(* IEC 61131-3 sources: plc-st-coding-agent/progress/evidence/f14_v14_remaining_20261113/jobs/codex_deepseek-v4pro, 118 files *)

(* ---- public-easy-01.candidate_01.st ---- *)
(*
ENGINEERING_CONTRACT
Pump_Motor: set by bottleSensor in Idle (PUB001), hold in Cleaning, reset by cleaningConfirmButton -> Filling (PUB002), BOOL.
Filling_Valve: set by cleaningConfirmButton in Cleaning (PUB002), hold in Filling, reset by fillingConfirmButton -> Capping (PUB003), BOOL.
Capping_Machine: set by fillingConfirmButton in Filling (PUB003), hold in Capping, reset by cappingConfirmButton -> Packing (PUB004), BOOL.
Packing_Machine: set by cappingConfirmButton in Capping (PUB004), hold in Packing, reset by packingConfirmButton -> Completed (PUB005), BOOL.
Completion_Light: set by packingConfirmButton in Packing (PUB005), hold in Completed, reset by finishedButton -> Idle (PUB006), BOOL.
Same-scan: one state transition per scan from the current state; later inputs are processed on subsequent scans. No numeric boundaries.
*)

(* CONTRACT_RULES [{"kind":"hold_until_reset","output":"Pump_Motor","set_input":"bottleSensor","reset_input":"cleaningConfirmButton"},{"kind":"hold_until_reset","output":"Filling_Valve","set_input":"cleaningConfirmButton","reset_input":"fillingConfirmButton"},{"kind":"hold_until_reset","output":"Capping_Machine","set_input":"fillingConfirmButton","reset_input":"cappingConfirmButton"},{"kind":"hold_until_reset","output":"Packing_Machine","set_input":"cappingConfirmButton","reset_input":"packingConfirmButton"},{"kind":"hold_until_reset","output":"Completion_Light","set_input":"packingConfirmButton","reset_input":"finishedButton"}] *)

FUNCTION_BLOCK FillingLineControl
VAR_INPUT
    bottleSensor : BOOL;
    cleaningConfirmButton : BOOL;
    fillingConfirmButton : BOOL;
    cappingConfirmButton : BOOL;
    packingConfirmButton : BOOL;
    finishedButton : BOOL;
END_VAR
VAR_OUTPUT
    Pump_Motor : BOOL;
    Filling_Valve : BOOL;
    Capping_Machine : BOOL;
    Packing_Machine : BOOL;
    Completion_Light : BOOL;
END_VAR
VAR
    State : INT := 0;
END_VAR

IF State = 0 AND bottleSensor THEN
    State := 1;
ELSIF State = 1 AND cleaningConfirmButton THEN
    State := 2;
ELSIF State = 2 AND fillingConfirmButton THEN
    State := 3;
ELSIF State = 3 AND cappingConfirmButton THEN
    State := 4;
ELSIF State = 4 AND packingConfirmButton THEN
    State := 5;
ELSIF State = 5 AND finishedButton THEN
    State := 0;
END_IF;

Pump_Motor := (State = 1);
Filling_Valve := (State = 2);
Capping_Machine := (State = 3);
Packing_Machine := (State = 4);
Completion_Light := (State = 5);

END_FUNCTION_BLOCK

(* ---- public-easy-01.candidate_02.st ---- *)
(*
ENGINEERING_CONTRACT
Pump_Motor: set by bottleSensor; retained until finishedButton resets the cycle. BOOL output.
Filling_Valve: set by cleaningConfirmButton; retained until finishedButton resets the cycle. BOOL output.
Capping_Machine: set by fillingConfirmButton; retained until finishedButton resets the cycle. BOOL output.
Packing_Machine: set by cappingConfirmButton; retained until finishedButton resets the cycle. BOOL output.
Completion_Light: set by packingConfirmButton; reset by finishedButton (PUB006). BOOL output.
Later stage confirmations are not explicit stop events, so earlier outputs remain active. No numeric boundaries.
Same-scan: finishedButton reset takes priority over activation inputs.
*)

(* CONTRACT_RULES [{"kind":"hold_until_reset","output":"Pump_Motor","set_input":"bottleSensor","reset_input":"finishedButton"},{"kind":"hold_until_reset","output":"Filling_Valve","set_input":"cleaningConfirmButton","reset_input":"finishedButton"},{"kind":"hold_until_reset","output":"Capping_Machine","set_input":"fillingConfirmButton","reset_input":"finishedButton"},{"kind":"hold_until_reset","output":"Packing_Machine","set_input":"cappingConfirmButton","reset_input":"finishedButton"},{"kind":"hold_until_reset","output":"Completion_Light","set_input":"packingConfirmButton","reset_input":"finishedButton"}] *)

FUNCTION_BLOCK FillingLineControl
VAR_INPUT
    bottleSensor : BOOL;
    cleaningConfirmButton : BOOL;
    fillingConfirmButton : BOOL;
    cappingConfirmButton : BOOL;
    packingConfirmButton : BOOL;
    finishedButton : BOOL;
END_VAR
VAR_OUTPUT
    Pump_Motor : BOOL;
    Filling_Valve : BOOL;
    Capping_Machine : BOOL;
    Packing_Machine : BOOL;
    Completion_Light : BOOL;
END_VAR
IF finishedButton THEN
    Pump_Motor := FALSE;
    Filling_Valve := FALSE;
    Capping_Machine := FALSE;
    Packing_Machine := FALSE;
    Completion_Light := FALSE;
ELSE
    IF bottleSensor THEN
        Pump_Motor := TRUE;
    END_IF;
    IF cleaningConfirmButton THEN
        Filling_Valve := TRUE;
    END_IF;
    IF fillingConfirmButton THEN
        Capping_Machine := TRUE;
    END_IF;
    IF cappingConfirmButton THEN
        Packing_Machine := TRUE;
    END_IF;
    IF packingConfirmButton THEN
        Completion_Light := TRUE;
    END_IF;
END_IF;

END_FUNCTION_BLOCK

(* ---- public-easy-01.candidate_03.st ---- *)
(*
ENGINEERING_CONTRACT
Pump_Motor: set by bottleSensor; retained until finishedButton resets the cycle. BOOL output.
Filling_Valve: set by cleaningConfirmButton; retained until finishedButton resets the cycle. BOOL output.
Capping_Machine: set by fillingConfirmButton; retained until finishedButton resets the cycle. BOOL output.
Packing_Machine: set by cappingConfirmButton while Capping_Machine is active; retained until finishedButton resets the cycle. BOOL output.
Completion_Light: set by packingConfirmButton while Packing_Machine is active; reset by finishedButton (PUB006). BOOL output.
Later stage confirmations are not explicit stop events, so earlier outputs remain active. No numeric boundaries.
Same-scan: finishedButton reset takes priority over activation inputs.
*)

(* CONTRACT_RULES [{"kind":"hold_until_reset","output":"Pump_Motor","set_input":"bottleSensor","reset_input":"finishedButton"}] *)

FUNCTION_BLOCK FillingLineControl
VAR_INPUT
    bottleSensor : BOOL;
    cleaningConfirmButton : BOOL;
    fillingConfirmButton : BOOL;
    cappingConfirmButton : BOOL;
    packingConfirmButton : BOOL;
    finishedButton : BOOL;
END_VAR
VAR_OUTPUT
    Pump_Motor : BOOL;
    Filling_Valve : BOOL;
    Capping_Machine : BOOL;
    Packing_Machine : BOOL;
    Completion_Light : BOOL;
END_VAR
IF finishedButton THEN
    Pump_Motor := FALSE;
    Filling_Valve := FALSE;
    Capping_Machine := FALSE;
    Packing_Machine := FALSE;
    Completion_Light := FALSE;
ELSE
    IF bottleSensor THEN
        Pump_Motor := TRUE;
    END_IF;
    IF cleaningConfirmButton THEN
        Filling_Valve := TRUE;
    END_IF;
    IF fillingConfirmButton THEN
        Capping_Machine := TRUE;
    END_IF;
    IF cappingConfirmButton AND Capping_Machine THEN
        Packing_Machine := TRUE;
    END_IF;
    IF packingConfirmButton AND Packing_Machine THEN
        Completion_Light := TRUE;
    END_IF;
END_IF;

END_FUNCTION_BLOCK

(* ---- public-easy-01.candidate_04.st ---- *)
(*
ENGINEERING_CONTRACT
Pump_Motor: set by bottleSensor; retained until finishedButton resets the cycle. BOOL output.
Filling_Valve: set by cleaningConfirmButton; retained until finishedButton resets the cycle. BOOL output.
Capping_Machine: set by fillingConfirmButton; retained until finishedButton resets the cycle. BOOL output.
Packing_Machine: set by cappingConfirmButton; retained until finishedButton resets the cycle. BOOL output.
Completion_Light: set by packingConfirmButton; reset by finishedButton (PUB006). BOOL output.
Later stage confirmations are not explicit stop events, so earlier outputs remain active. No numeric boundaries.
Same-scan: finishedButton reset takes priority over activation inputs.
*)

(* CONTRACT_RULES [{"kind":"hold_until_reset","output":"Pump_Motor","set_input":"bottleSensor","reset_input":"finishedButton"}] *)

FUNCTION_BLOCK FillingLineControl
VAR_INPUT
    bottleSensor : BOOL;
    cleaningConfirmButton : BOOL;
    fillingConfirmButton : BOOL;
    cappingConfirmButton : BOOL;
    packingConfirmButton : BOOL;
    finishedButton : BOOL;
END_VAR
VAR_OUTPUT
    Pump_Motor : BOOL;
    Filling_Valve : BOOL;
    Capping_Machine : BOOL;
    Packing_Machine : BOOL;
    Completion_Light : BOOL;
END_VAR
IF finishedButton THEN
    Pump_Motor := FALSE;
    Filling_Valve := FALSE;
    Capping_Machine := FALSE;
    Packing_Machine := FALSE;
    Completion_Light := FALSE;
ELSE
    IF bottleSensor THEN
        Pump_Motor := TRUE;
    END_IF;
    IF cleaningConfirmButton THEN
        Filling_Valve := TRUE;
    END_IF;
    IF fillingConfirmButton THEN
        Capping_Machine := TRUE;
    END_IF;
    IF cappingConfirmButton THEN
        Packing_Machine := TRUE;
    END_IF;
    IF packingConfirmButton THEN
        Completion_Light := TRUE;
    END_IF;
END_IF;

END_FUNCTION_BLOCK

(* ---- public-easy-01.patch_base_02.st ---- *)
(*
ENGINEERING_CONTRACT
Pump_Motor: set by bottleSensor in Idle (PUB001), hold in Cleaning, reset by cleaningConfirmButton -> Filling (PUB002), BOOL.
Filling_Valve: set by cleaningConfirmButton in Cleaning (PUB002), hold in Filling, reset by fillingConfirmButton -> Capping (PUB003), BOOL.
Capping_Machine: set by fillingConfirmButton in Filling (PUB003), hold in Capping, reset by cappingConfirmButton -> Packing (PUB004), BOOL.
Packing_Machine: set by cappingConfirmButton in Capping (PUB004), hold in Packing, reset by packingConfirmButton -> Completed (PUB005), BOOL.
Completion_Light: set by packingConfirmButton in Packing (PUB005), hold in Completed, reset by finishedButton -> Idle (PUB006), BOOL.
Same-scan: one state transition per scan from the current state; later inputs are processed on subsequent scans. No numeric boundaries.
*)

(* CONTRACT_RULES [{"kind":"hold_until_reset","output":"Pump_Motor","set_input":"bottleSensor","reset_input":"cleaningConfirmButton"},{"kind":"hold_until_reset","output":"Filling_Valve","set_input":"cleaningConfirmButton","reset_input":"fillingConfirmButton"},{"kind":"hold_until_reset","output":"Capping_Machine","set_input":"fillingConfirmButton","reset_input":"cappingConfirmButton"},{"kind":"hold_until_reset","output":"Packing_Machine","set_input":"cappingConfirmButton","reset_input":"packingConfirmButton"},{"kind":"hold_until_reset","output":"Completion_Light","set_input":"packingConfirmButton","reset_input":"finishedButton"}] *)

FUNCTION_BLOCK FillingLineControl
VAR_INPUT
    bottleSensor : BOOL;
    cleaningConfirmButton : BOOL;
    fillingConfirmButton : BOOL;
    cappingConfirmButton : BOOL;
    packingConfirmButton : BOOL;
    finishedButton : BOOL;
END_VAR
VAR_OUTPUT
    Pump_Motor : BOOL;
    Filling_Valve : BOOL;
    Capping_Machine : BOOL;
    Packing_Machine : BOOL;
    Completion_Light : BOOL;
END_VAR
VAR
    State : INT := 0;
END_VAR

IF State = 0 AND bottleSensor THEN
    State := 1;
ELSIF State = 1 AND cleaningConfirmButton THEN
    State := 2;
ELSIF State = 2 AND fillingConfirmButton THEN
    State := 3;
ELSIF State = 3 AND cappingConfirmButton THEN
    State := 4;
ELSIF State = 4 AND packingConfirmButton THEN
    State := 5;
ELSIF State = 5 AND finishedButton THEN
    State := 0;
END_IF;

Pump_Motor := (State = 1);
Filling_Valve := (State = 2);
Capping_Machine := (State = 3);
Packing_Machine := (State = 4);
Completion_Light := (State = 5);

END_FUNCTION_BLOCK

(* ---- public-easy-01.patch_base_03.st ---- *)
(*
ENGINEERING_CONTRACT
Pump_Motor: set by bottleSensor; retained until finishedButton resets the cycle. BOOL output.
Filling_Valve: set by cleaningConfirmButton; retained until finishedButton resets the cycle. BOOL output.
Capping_Machine: set by fillingConfirmButton; retained until finishedButton resets the cycle. BOOL output.
Packing_Machine: set by cappingConfirmButton; retained until finishedButton resets the cycle. BOOL output.
Completion_Light: set by packingConfirmButton; reset by finishedButton (PUB006). BOOL output.
Later stage confirmations are not explicit stop events, so earlier outputs remain active. No numeric boundaries.
Same-scan: finishedButton reset takes priority over activation inputs.
*)

(* CONTRACT_RULES [{"kind":"hold_until_reset","output":"Pump_Motor","set_input":"bottleSensor","reset_input":"finishedButton"},{"kind":"hold_until_reset","output":"Filling_Valve","set_input":"cleaningConfirmButton","reset_input":"finishedButton"},{"kind":"hold_until_reset","output":"Capping_Machine","set_input":"fillingConfirmButton","reset_input":"finishedButton"},{"kind":"hold_until_reset","output":"Packing_Machine","set_input":"cappingConfirmButton","reset_input":"finishedButton"},{"kind":"hold_until_reset","output":"Completion_Light","set_input":"packingConfirmButton","reset_input":"finishedButton"}] *)

FUNCTION_BLOCK FillingLineControl
VAR_INPUT
    bottleSensor : BOOL;
    cleaningConfirmButton : BOOL;
    fillingConfirmButton : BOOL;
    cappingConfirmButton : BOOL;
    packingConfirmButton : BOOL;
    finishedButton : BOOL;
END_VAR
VAR_OUTPUT
    Pump_Motor : BOOL;
    Filling_Valve : BOOL;
    Capping_Machine : BOOL;
    Packing_Machine : BOOL;
    Completion_Light : BOOL;
END_VAR
IF finishedButton THEN
    Pump_Motor := FALSE;
    Filling_Valve := FALSE;
    Capping_Machine := FALSE;
    Packing_Machine := FALSE;
    Completion_Light := FALSE;
ELSE
    IF bottleSensor THEN
        Pump_Motor := TRUE;
    END_IF;
    IF cleaningConfirmButton THEN
        Filling_Valve := TRUE;
    END_IF;
    IF fillingConfirmButton THEN
        Capping_Machine := TRUE;
    END_IF;
    IF cappingConfirmButton THEN
        Packing_Machine := TRUE;
    END_IF;
    IF packingConfirmButton THEN
        Completion_Light := TRUE;
    END_IF;
END_IF;

END_FUNCTION_BLOCK

(* ---- public-easy-01.patch_base_04.st ---- *)
(*
ENGINEERING_CONTRACT
Pump_Motor: set by bottleSensor; retained until finishedButton resets the cycle. BOOL output.
Filling_Valve: set by cleaningConfirmButton; retained until finishedButton resets the cycle. BOOL output.
Capping_Machine: set by fillingConfirmButton; retained until finishedButton resets the cycle. BOOL output.
Packing_Machine: set by cappingConfirmButton while Capping_Machine is active; retained until finishedButton resets the cycle. BOOL output.
Completion_Light: set by packingConfirmButton while Packing_Machine is active; reset by finishedButton (PUB006). BOOL output.
Later stage confirmations are not explicit stop events, so earlier outputs remain active. No numeric boundaries.
Same-scan: finishedButton reset takes priority over activation inputs.
*)

(* CONTRACT_RULES [{"kind":"hold_until_reset","output":"Pump_Motor","set_input":"bottleSensor","reset_input":"finishedButton"}] *)

FUNCTION_BLOCK FillingLineControl
VAR_INPUT
    bottleSensor : BOOL;
    cleaningConfirmButton : BOOL;
    fillingConfirmButton : BOOL;
    cappingConfirmButton : BOOL;
    packingConfirmButton : BOOL;
    finishedButton : BOOL;
END_VAR
VAR_OUTPUT
    Pump_Motor : BOOL;
    Filling_Valve : BOOL;
    Capping_Machine : BOOL;
    Packing_Machine : BOOL;
    Completion_Light : BOOL;
END_VAR
IF finishedButton THEN
    Pump_Motor := FALSE;
    Filling_Valve := FALSE;
    Capping_Machine := FALSE;
    Packing_Machine := FALSE;
    Completion_Light := FALSE;
ELSE
    IF bottleSensor THEN
        Pump_Motor := TRUE;
    END_IF;
    IF cleaningConfirmButton THEN
        Filling_Valve := TRUE;
    END_IF;
    IF fillingConfirmButton THEN
        Capping_Machine := TRUE;
    END_IF;
    IF cappingConfirmButton AND Capping_Machine THEN
        Packing_Machine := TRUE;
    END_IF;
    IF packingConfirmButton AND Packing_Machine THEN
        Completion_Light := TRUE;
    END_IF;
END_IF;

END_FUNCTION_BLOCK

(* ---- public-easy-01.raw_candidate_01.st ---- *)
(*
ENGINEERING_CONTRACT
Pump_Motor: set by bottleSensor in Idle (PUB001), hold in Cleaning, reset by cleaningConfirmButton -> Filling (PUB002), BOOL.
Filling_Valve: set by cleaningConfirmButton in Cleaning (PUB002), hold in Filling, reset by fillingConfirmButton -> Capping (PUB003), BOOL.
Capping_Machine: set by fillingConfirmButton in Filling (PUB003), hold in Capping, reset by cappingConfirmButton -> Packing (PUB004), BOOL.
Packing_Machine: set by cappingConfirmButton in Capping (PUB004), hold in Packing, reset by packingConfirmButton -> Completed (PUB005), BOOL.
Completion_Light: set by packingConfirmButton in Packing (PUB005), hold in Completed, reset by finishedButton -> Idle (PUB006), BOOL.
Same-scan: one state transition per scan from the current state; later inputs are processed on subsequent scans. No numeric boundaries.
*)

(* CONTRACT_RULES [{"kind":"hold_until_reset","output":"Pump_Motor","set_input":"bottleSensor","reset_input":"cleaningConfirmButton"},{"kind":"hold_until_reset","output":"Filling_Valve","set_input":"cleaningConfirmButton","reset_input":"fillingConfirmButton"},{"kind":"hold_until_reset","output":"Capping_Machine","set_input":"fillingConfirmButton","reset_input":"cappingConfirmButton"},{"kind":"hold_until_reset","output":"Packing_Machine","set_input":"cappingConfirmButton","reset_input":"packingConfirmButton"},{"kind":"hold_until_reset","output":"Completion_Light","set_input":"packingConfirmButton","reset_input":"finishedButton"}] *)

FUNCTION_BLOCK FillingLineControl
VAR_INPUT
    bottleSensor : BOOL;
    cleaningConfirmButton : BOOL;
    fillingConfirmButton : BOOL;
    cappingConfirmButton : BOOL;
    packingConfirmButton : BOOL;
    finishedButton : BOOL;
END_VAR
VAR_OUTPUT
    Pump_Motor : BOOL;
    Filling_Valve : BOOL;
    Capping_Machine : BOOL;
    Packing_Machine : BOOL;
    Completion_Light : BOOL;
END_VAR
VAR
    State : INT := 0;
END_VAR

IF State = 0 AND bottleSensor THEN
    State := 1;
ELSIF State = 1 AND cleaningConfirmButton THEN
    State := 2;
ELSIF State = 2 AND fillingConfirmButton THEN
    State := 3;
ELSIF State = 3 AND cappingConfirmButton THEN
    State := 4;
ELSIF State = 4 AND packingConfirmButton THEN
    State := 5;
ELSIF State = 5 AND finishedButton THEN
    State := 0;
END_IF;

Pump_Motor := (State = 1);
Filling_Valve := (State = 2);
Capping_Machine := (State = 3);
Packing_Machine := (State = 4);
Completion_Light := (State = 5);

END_FUNCTION_BLOCK

(* ---- public-easy-01.raw_candidate_02.st ---- *)
(*
ENGINEERING_CONTRACT
Pump_Motor: set by bottleSensor; retained until finishedButton resets the cycle. BOOL output.
Filling_Valve: set by cleaningConfirmButton; retained until finishedButton resets the cycle. BOOL output.
Capping_Machine: set by fillingConfirmButton; retained until finishedButton resets the cycle. BOOL output.
Packing_Machine: set by cappingConfirmButton; retained until finishedButton resets the cycle. BOOL output.
Completion_Light: set by packingConfirmButton; reset by finishedButton (PUB006). BOOL output.
Later stage confirmations are not explicit stop events, so earlier outputs remain active. No numeric boundaries.
Same-scan: finishedButton reset takes priority over activation inputs.
*)

(* CONTRACT_RULES [{"kind":"hold_until_reset","output":"Pump_Motor","set_input":"bottleSensor","reset_input":"finishedButton"},{"kind":"hold_until_reset","output":"Filling_Valve","set_input":"cleaningConfirmButton","reset_input":"finishedButton"},{"kind":"hold_until_reset","output":"Capping_Machine","set_input":"fillingConfirmButton","reset_input":"finishedButton"},{"kind":"hold_until_reset","output":"Packing_Machine","set_input":"cappingConfirmButton","reset_input":"finishedButton"},{"kind":"hold_until_reset","output":"Completion_Light","set_input":"packingConfirmButton","reset_input":"finishedButton"}] *)

FUNCTION_BLOCK FillingLineControl
VAR_INPUT
    bottleSensor : BOOL;
    cleaningConfirmButton : BOOL;
    fillingConfirmButton : BOOL;
    cappingConfirmButton : BOOL;
    packingConfirmButton : BOOL;
    finishedButton : BOOL;
END_VAR
VAR_OUTPUT
    Pump_Motor : BOOL;
    Filling_Valve : BOOL;
    Capping_Machine : BOOL;
    Packing_Machine : BOOL;
    Completion_Light : BOOL;
END_VAR
IF finishedButton THEN
    Pump_Motor := FALSE;
    Filling_Valve := FALSE;
    Capping_Machine := FALSE;
    Packing_Machine := FALSE;
    Completion_Light := FALSE;
ELSE
    IF bottleSensor THEN
        Pump_Motor := TRUE;
    END_IF;
    IF cleaningConfirmButton THEN
        Filling_Valve := TRUE;
    END_IF;
    IF fillingConfirmButton THEN
        Capping_Machine := TRUE;
    END_IF;
    IF cappingConfirmButton THEN
        Packing_Machine := TRUE;
    END_IF;
    IF packingConfirmButton THEN
        Completion_Light := TRUE;
    END_IF;
END_IF;

END_FUNCTION_BLOCK

(* ---- public-easy-01.raw_candidate_03.st ---- *)
(*
ENGINEERING_CONTRACT
Pump_Motor: set by bottleSensor; retained until finishedButton resets the cycle. BOOL output.
Filling_Valve: set by cleaningConfirmButton; retained until finishedButton resets the cycle. BOOL output.
Capping_Machine: set by fillingConfirmButton; retained until finishedButton resets the cycle. BOOL output.
Packing_Machine: set by cappingConfirmButton while Capping_Machine is active; retained until finishedButton resets the cycle. BOOL output.
Completion_Light: set by packingConfirmButton while Packing_Machine is active; reset by finishedButton (PUB006). BOOL output.
Later stage confirmations are not explicit stop events, so earlier outputs remain active. No numeric boundaries.
Same-scan: finishedButton reset takes priority over activation inputs.
*)

(* CONTRACT_RULES [{"kind":"hold_until_reset","output":"Pump_Motor","set_input":"bottleSensor","reset_input":"finishedButton"}] *)

FUNCTION_BLOCK FillingLineControl
VAR_INPUT
    bottleSensor : BOOL;
    cleaningConfirmButton : BOOL;
    fillingConfirmButton : BOOL;
    cappingConfirmButton : BOOL;
    packingConfirmButton : BOOL;
    finishedButton : BOOL;
END_VAR
VAR_OUTPUT
    Pump_Motor : BOOL;
    Filling_Valve : BOOL;
    Capping_Machine : BOOL;
    Packing_Machine : BOOL;
    Completion_Light : BOOL;
END_VAR
IF finishedButton THEN
    Pump_Motor := FALSE;
    Filling_Valve := FALSE;
    Capping_Machine := FALSE;
    Packing_Machine := FALSE;
    Completion_Light := FALSE;
ELSE
    IF bottleSensor THEN
        Pump_Motor := TRUE;
    END_IF;
    IF cleaningConfirmButton THEN
        Filling_Valve := TRUE;
    END_IF;
    IF fillingConfirmButton THEN
        Capping_Machine := TRUE;
    END_IF;
    IF cappingConfirmButton AND Capping_Machine THEN
        Packing_Machine := TRUE;
    END_IF;
    IF packingConfirmButton AND Packing_Machine THEN
        Completion_Light := TRUE;
    END_IF;
END_IF;

END_FUNCTION_BLOCK

(* ---- public-easy-01.raw_candidate_04.st ---- *)
(*
ENGINEERING_CONTRACT
Pump_Motor: set by bottleSensor; retained until finishedButton resets the cycle. BOOL output.
Filling_Valve: set by cleaningConfirmButton; retained until finishedButton resets the cycle. BOOL output.
Capping_Machine: set by fillingConfirmButton; retained until finishedButton resets the cycle. BOOL output.
Packing_Machine: set by cappingConfirmButton; retained until finishedButton resets the cycle. BOOL output.
Completion_Light: set by packingConfirmButton; reset by finishedButton (PUB006). BOOL output.
Later stage confirmations are not explicit stop events, so earlier outputs remain active. No numeric boundaries.
Same-scan: finishedButton reset takes priority over activation inputs.
*)

(* CONTRACT_RULES [{"kind":"hold_until_reset","output":"Pump_Motor","set_input":"bottleSensor","reset_input":"finishedButton"}] *)

FUNCTION_BLOCK FillingLineControl
VAR_INPUT
    bottleSensor : BOOL;
    cleaningConfirmButton : BOOL;
    fillingConfirmButton : BOOL;
    cappingConfirmButton : BOOL;
    packingConfirmButton : BOOL;
    finishedButton : BOOL;
END_VAR
VAR_OUTPUT
    Pump_Motor : BOOL;
    Filling_Valve : BOOL;
    Capping_Machine : BOOL;
    Packing_Machine : BOOL;
    Completion_Light : BOOL;
END_VAR
IF finishedButton THEN
    Pump_Motor := FALSE;
    Filling_Valve := FALSE;
    Capping_Machine := FALSE;
    Packing_Machine := FALSE;
    Completion_Light := FALSE;
ELSE
    IF bottleSensor THEN
        Pump_Motor := TRUE;
    END_IF;
    IF cleaningConfirmButton THEN
        Filling_Valve := TRUE;
    END_IF;
    IF fillingConfirmButton THEN
        Capping_Machine := TRUE;
    END_IF;
    IF cappingConfirmButton THEN
        Packing_Machine := TRUE;
    END_IF;
    IF packingConfirmButton THEN
        Completion_Light := TRUE;
    END_IF;
END_IF;

END_FUNCTION_BLOCK

(* ---- public-easy-02.candidate_01.st ---- *)
(*
ENGINEERING_CONTRACT
- Scope: PUB001, DWORD edge detection reported every scan.
- hasChanged: combinational; TRUE when current value differs from previous scan.
- risingBits/fallingBits: current-scan edge masks, recomputed every call; no retention.
- hasRisingEdges/hasFallingEdges: combinational nonzero-mask indicators.
- noOfRisingBits/noOfFallingBits: USINT popcount, 0..32, unit = edge count.
- State update: previous value stored after outputs are evaluated.
- First-scan baseline: unspecified; implemented as zero-initialized previous value.
- Same-scan priority: edges are functions of the current value and the prior value.
*)

(* CONTRACT_RULES [] *)

FUNCTION_BLOCK FB
VAR_INPUT
    value : DWORD;
END_VAR
VAR_OUTPUT
    hasChanged : BOOL;
    hasRisingEdges : BOOL;
    risingBits : DWORD;
    noOfRisingBits : USINT;
    hasFallingEdges : BOOL;
    fallingBits : DWORD;
    noOfFallingBits : USINT;
END_VAR
VAR
    local_lastValue : DWORD := DWORD#0;
    tmp_bitIndex : INT;
    tmp_bitMask : DWORD;
END_VAR

hasChanged := value <> local_lastValue;
risingBits := (NOT local_lastValue) AND value;
fallingBits := local_lastValue AND (NOT value);

hasRisingEdges := risingBits <> DWORD#0;
hasFallingEdges := fallingBits <> DWORD#0;

noOfRisingBits := 0;
noOfFallingBits := 0;

FOR tmp_bitIndex := 0 TO 31 DO
    tmp_bitMask := SHL(DWORD#1, tmp_bitIndex);
    IF (risingBits AND tmp_bitMask) <> DWORD#0 THEN
        noOfRisingBits := noOfRisingBits + 1;
    END_IF;
    IF (fallingBits AND tmp_bitMask) <> DWORD#0 THEN
        noOfFallingBits := noOfFallingBits + 1;
    END_IF;
END_FOR;

local_lastValue := value;
END_FUNCTION_BLOCK

(* ---- public-easy-02.raw_candidate_01.st ---- *)
(*
ENGINEERING_CONTRACT
- Scope: PUB001, DWORD edge detection reported every scan.
- hasChanged: combinational; TRUE when current value differs from previous scan.
- risingBits/fallingBits: current-scan edge masks, recomputed every call; no retention.
- hasRisingEdges/hasFallingEdges: combinational nonzero-mask indicators.
- noOfRisingBits/noOfFallingBits: USINT popcount, 0..32, unit = edge count.
- State update: previous value stored after outputs are evaluated.
- First-scan baseline: unspecified; implemented as zero-initialized previous value.
- Same-scan priority: edges are functions of the current value and the prior value.
*)

(* CONTRACT_RULES [] *)

FUNCTION_BLOCK FB
VAR_INPUT
    value : DWORD;
END_VAR
VAR_OUTPUT
    hasChanged : BOOL;
    hasRisingEdges : BOOL;
    risingBits : DWORD;
    noOfRisingBits : USINT;
    hasFallingEdges : BOOL;
    fallingBits : DWORD;
    noOfFallingBits : USINT;
END_VAR
VAR
    local_lastValue : DWORD := DWORD#0;
    tmp_bitIndex : INT;
    tmp_bitMask : DWORD;
END_VAR

hasChanged := value <> local_lastValue;
risingBits := (NOT local_lastValue) AND value;
fallingBits := local_lastValue AND (NOT value);

hasRisingEdges := risingBits <> DWORD#0;
hasFallingEdges := fallingBits <> DWORD#0;

noOfRisingBits := 0;
noOfFallingBits := 0;

FOR tmp_bitIndex := 0 TO 31 DO
    tmp_bitMask := SHL(DWORD#1, tmp_bitIndex);
    IF (risingBits AND tmp_bitMask) <> DWORD#0 THEN
        noOfRisingBits := noOfRisingBits + 1;
    END_IF;
    IF (fallingBits AND tmp_bitMask) <> DWORD#0 THEN
        noOfFallingBits := noOfFallingBits + 1;
    END_IF;
END_FOR;

local_lastValue := value;
END_FUNCTION_BLOCK

(* ---- public-easy-03.candidate_01.st ---- *)
FUNCTION_BLOCK AlarmHandling
VAR_INPUT
    Value : REAL;
    hiLevel : REAL;
    loLevel : REAL;
    hystWindow : REAL;
END_VAR
VAR_OUTPUT
    hiAlarm : BOOL;
    loAlarm : BOOL;
    error : BOOL;
    status : WORD;
END_VAR
VAR
END_VAR

(* ENGINEERING_CONTRACT
  hiAlarm: set while Value > hiLevel (PUB001); retained until Value < hiLevel-hystWindow (PUB001/PUB002).
  loAlarm: set while Value < loLevel (PUB001); retained until Value > loLevel+hystWindow (PUB001/PUB002).
  error/16#8001: loLevel >= hiLevel has priority, returns immediately after setting error and clearing alarms (PUB003).
  error/16#8002: hystWindow >= hiLevel-loLevel returns immediately after setting error and clearing alarms (PUB004).
  valid configuration: error := FALSE, status := 0, then both alarm paths are evaluated in the same scan.
  strict > and < comparisons only; equality retains the current alarm state. REAL boundaries and thresholds.
*)

(* CONTRACT_RULES [] *)

IF loLevel >= hiLevel THEN
    error := TRUE;
    status := 16#8001;
    hiAlarm := FALSE;
    loAlarm := FALSE;
    RETURN;
END_IF;

IF hystWindow >= hiLevel - loLevel THEN
    error := TRUE;
    status := 16#8002;
    hiAlarm := FALSE;
    loAlarm := FALSE;
    RETURN;
END_IF;

error := FALSE;
status := 0;

IF Value > hiLevel THEN
    hiAlarm := TRUE;
ELSIF Value < hiLevel - hystWindow THEN
    hiAlarm := FALSE;
END_IF;

IF Value < loLevel THEN
    loAlarm := TRUE;
ELSIF Value > loLevel + hystWindow THEN
    loAlarm := FALSE;
END_IF;

END_FUNCTION_BLOCK

(* ---- public-easy-03.raw_candidate_01.st ---- *)
FUNCTION_BLOCK AlarmHandling
VAR_INPUT
    Value : REAL;
    hiLevel : REAL;
    loLevel : REAL;
    hystWindow : REAL;
END_VAR
VAR_OUTPUT
    hiAlarm : BOOL;
    loAlarm : BOOL;
    error : BOOL;
    status : WORD;
END_VAR
VAR
END_VAR

(* ENGINEERING_CONTRACT
  hiAlarm: set while Value > hiLevel (PUB001); retained until Value < hiLevel-hystWindow (PUB001/PUB002).
  loAlarm: set while Value < loLevel (PUB001); retained until Value > loLevel+hystWindow (PUB001/PUB002).
  error/16#8001: loLevel >= hiLevel has priority, returns immediately after setting error and clearing alarms (PUB003).
  error/16#8002: hystWindow >= hiLevel-loLevel returns immediately after setting error and clearing alarms (PUB004).
  valid configuration: error := FALSE, status := 0, then both alarm paths are evaluated in the same scan.
  strict > and < comparisons only; equality retains the current alarm state. REAL boundaries and thresholds.
*)

(* CONTRACT_RULES [] *)

IF loLevel >= hiLevel THEN
    error := TRUE;
    status := 16#8001;
    hiAlarm := FALSE;
    loAlarm := FALSE;
    RETURN;
END_IF

IF hystWindow >= hiLevel - loLevel THEN
    error := TRUE;
    status := 16#8002;
    hiAlarm := FALSE;
    loAlarm := FALSE;
    RETURN;
END_IF

error := FALSE;
status := 0;

IF Value > hiLevel THEN
    hiAlarm := TRUE;
ELSIF Value < hiLevel - hystWindow THEN
    hiAlarm := FALSE;
END_IF

IF Value < loLevel THEN
    loAlarm := TRUE;
ELSIF Value > loLevel + hystWindow THEN
    loAlarm := FALSE;
END_IF

END_FUNCTION_BLOCK

(* ---- public-easy-04.candidate_01.st ---- *)
FUNCTION_BLOCK FB_JamPumpControl
VAR_INPUT
    VISCOSITY_OK : BOOL;
    PASTE_E_STOP_NC : BOOL;
    DebounceTime : TIME;
    CycleTime : TIME;
END_VAR
VAR_OUTPUT
    VFD_RUN : BOOL;
    PUMP_MAINT_DUE : BOOL;
    PUMP_RUNTIME_ACC : LTIME;
END_VAR
VAR
    tmp_first_scan : BOOL := TRUE;
    tmp_debounce_enable : BOOL;
    tmp_debounce_timer : TON;
    tmp_viscosity_valid : BOOL;
    tmp_runtime_acc : LTIME;
    tmp_maintenance_threshold : LTIME;
END_VAR

(* ENGINEERING_CONTRACT
VFD_RUN: active iff PASTE_E_STOP_NC AND tmp_viscosity_valid; any false permissive deactivates immediately; final same-scan inputs decide run and accumulation (PUB002).
Debounce validity: set same scan TON.Q fires; hold while VISCOSITY_OK remains TRUE; reset only when VISCOSITY_OK=FALSE (PUB001).
E-stop: clears incomplete debounce timing; completed viscosity validity is retained while VISCOSITY_OK remains TRUE (PUB002).
PUMP_RUNTIME_ACC: add TIME_TO_LTIME(CycleTime) only when final VFD_RUN=TRUE; preserve while stopped; starts at 0ns (PUB003).
PUMP_MAINT_DUE: remains TRUE when accumulated LTIME >= TIME_TO_LTIME(T#500h); informational only; starts FALSE (PUB004).
Initialization: first scan sets run OFF, accumulated runtime 0ns, maintenance FALSE (PUB005).
Units: TIME inputs in ms; LTIME accumulation in ns; maintenance threshold strictly by >= at 500h.
*)

(* CONTRACT_RULES [] *)

IF tmp_first_scan THEN
    tmp_first_scan := FALSE;
    tmp_viscosity_valid := FALSE;
    tmp_runtime_acc := TIME_TO_LTIME(T#0ms);
    VFD_RUN := FALSE;
    PUMP_MAINT_DUE := FALSE;
    PUMP_RUNTIME_ACC := TIME_TO_LTIME(T#0ms);
END_IF;

tmp_maintenance_threshold := TIME_TO_LTIME(T#500h);
tmp_debounce_enable := VISCOSITY_OK AND PASTE_E_STOP_NC AND NOT tmp_viscosity_valid;
tmp_debounce_timer(IN := tmp_debounce_enable, PT := DebounceTime);

IF VISCOSITY_OK THEN
    IF tmp_debounce_timer.Q THEN
        tmp_viscosity_valid := TRUE;
    END_IF;
ELSE
    tmp_viscosity_valid := FALSE;
END_IF;

VFD_RUN := PASTE_E_STOP_NC AND tmp_viscosity_valid;

IF VFD_RUN THEN
    tmp_runtime_acc := tmp_runtime_acc + TIME_TO_LTIME(CycleTime);
END_IF;

PUMP_RUNTIME_ACC := tmp_runtime_acc;
PUMP_MAINT_DUE := tmp_runtime_acc >= tmp_maintenance_threshold;

END_FUNCTION_BLOCK

(* ---- public-easy-04.raw_candidate_01.st ---- *)
FUNCTION_BLOCK FB_JamPumpControl
VAR_INPUT
    VISCOSITY_OK : BOOL;
    PASTE_E_STOP_NC : BOOL;
    DebounceTime : TIME;
    CycleTime : TIME;
END_VAR
VAR_OUTPUT
    VFD_RUN : BOOL;
    PUMP_MAINT_DUE : BOOL;
    PUMP_RUNTIME_ACC : LTIME;
END_VAR
VAR
    tmp_first_scan : BOOL := TRUE;
    tmp_debounce_enable : BOOL;
    tmp_debounce_timer : TON;
    tmp_viscosity_valid : BOOL;
    tmp_runtime_acc : LTIME;
    tmp_maintenance_threshold : LTIME;
END_VAR

(* ENGINEERING_CONTRACT
VFD_RUN: active iff PASTE_E_STOP_NC AND tmp_viscosity_valid; any false permissive deactivates immediately; final same-scan inputs decide run and accumulation (PUB002).
Debounce validity: set same scan TON.Q fires; hold while VISCOSITY_OK remains TRUE; reset only when VISCOSITY_OK=FALSE (PUB001).
E-stop: clears incomplete debounce timing; completed viscosity validity is retained while VISCOSITY_OK remains TRUE (PUB002).
PUMP_RUNTIME_ACC: add TIME_TO_LTIME(CycleTime) only when final VFD_RUN=TRUE; preserve while stopped; starts at 0ns (PUB003).
PUMP_MAINT_DUE: remains TRUE when accumulated LTIME >= TIME_TO_LTIME(T#500h); informational only; starts FALSE (PUB004).
Initialization: first scan sets run OFF, accumulated runtime 0ns, maintenance FALSE (PUB005).
Units: TIME inputs in ms; LTIME accumulation in ns; maintenance threshold strictly by >= at 500h.
*)

(* CONTRACT_RULES [] *)

IF tmp_first_scan THEN
    tmp_first_scan := FALSE;
    tmp_viscosity_valid := FALSE;
    tmp_runtime_acc := TIME_TO_LTIME(T#0ms);
    VFD_RUN := FALSE;
    PUMP_MAINT_DUE := FALSE;
    PUMP_RUNTIME_ACC := TIME_TO_LTIME(T#0ms);
END_IF;

tmp_maintenance_threshold := TIME_TO_LTIME(T#500h);
tmp_debounce_enable := VISCOSITY_OK AND PASTE_E_STOP_NC AND NOT tmp_viscosity_valid;
tmp_debounce_timer(IN := tmp_debounce_enable, PT := DebounceTime);

IF VISCOSITY_OK THEN
    IF tmp_debounce_timer.Q THEN
        tmp_viscosity_valid := TRUE;
    END_IF;
ELSE
    tmp_viscosity_valid := FALSE;
END_IF;

VFD_RUN := PASTE_E_STOP_NC AND tmp_viscosity_valid;

IF VFD_RUN THEN
    tmp_runtime_acc := tmp_runtime_acc + TIME_TO_LTIME(CycleTime);
END_IF;

PUMP_RUNTIME_ACC := tmp_runtime_acc;
PUMP_MAINT_DUE := tmp_runtime_acc >= tmp_maintenance_threshold;

END_FUNCTION_BLOCK

(* ---- public-easy-05.candidate_01.st ---- *)
FUNCTION_BLOCK WeldGapAlarm
VAR_INPUT
    Gap_Exceeded : BOOL;
    Weld_E_Stop_NC : BOOL;
    DebounceTime : TIME;
END_VAR
VAR_OUTPUT
    Operator_Alert : BOOL;
    Weld_Soft_Start_Active : BOOL;
END_VAR
VAR
    local_PowerUpTimer : TON;
    local_DebounceTimer : TON;
    local_DebounceEnable : BOOL;
END_VAR

(* CONTRACT_RULES [] *)

(* ENGINEERING_CONTRACT
Operator_Alert:
  Activate when E-stop inactive, power-up timer completed, and Gap_Exceeded has been TRUE continuously for DebounceTime.
  Hold while Gap_Exceeded remains TRUE after elapsed DebounceTime.
  Reset immediately on Gap_Exceeded=FALSE, E-stop active, or during initialization.
  Same-scan priority: E-stop active > initialization > debounced gap alarm.
Weld_Soft_Start_Active:
  Activate at power-up and hold TRUE for exactly the 5 s initialization period.
  Deactivate automatically when local_PowerUpTimer reaches 5 s; no manual reset.
  Same-scan priority: independent of E-stop and alarm deactivation.
Units/boundaries: power-up interval = T#5S; DebounceTime is TIME in milliseconds and must be positive.
*)

local_PowerUpTimer(IN := TRUE, PT := T#5S);

local_DebounceEnable := NOT local_PowerUpTimer.Q
                        AND Weld_E_Stop_NC
                        AND Gap_Exceeded;

local_DebounceTimer(IN := local_DebounceEnable, PT := DebounceTime);

Weld_Soft_Start_Active := NOT local_PowerUpTimer.Q;
Operator_Alert := Weld_E_Stop_NC AND local_DebounceTimer.Q;

END_FUNCTION_BLOCK

(* ---- public-easy-05.candidate_02.st ---- *)
FUNCTION_BLOCK WeldGapAlarm
VAR_INPUT
    Gap_Exceeded : BOOL;
    Weld_E_Stop_NC : BOOL;
    DebounceTime : TIME;
END_VAR
VAR_OUTPUT
    Operator_Alert : BOOL;
    Weld_Soft_Start_Active : BOOL;
END_VAR
VAR
    local_PowerUpTimer : TON;
    local_DebounceTimer : TON;
    local_DebounceEnable : BOOL;
END_VAR

(* CONTRACT_RULES [] *)

(* ENGINEERING_CONTRACT
Operator_Alert:
  Activate when E-stop inactive, power-up timer completed, and Gap_Exceeded has been TRUE continuously for DebounceTime.
  Hold while Gap_Exceeded remains TRUE after elapsed DebounceTime.
  Reset immediately on Gap_Exceeded=FALSE, E-stop active, or during initialization.
  Same-scan priority: E-stop active > initialization > debounced gap alarm.
Weld_Soft_Start_Active:
  Activate at power-up and hold TRUE for exactly the 5 s initialization period.
  Deactivate automatically when local_PowerUpTimer reaches 5 s; no manual reset.
  Same-scan priority: independent of E-stop and alarm deactivation.
Units/boundaries: power-up interval = T#5S; DebounceTime is TIME in milliseconds and must be positive.
*)

local_PowerUpTimer(IN := TRUE, PT := T#5S);

local_DebounceEnable := local_PowerUpTimer.Q
                        AND Weld_E_Stop_NC
                        AND Gap_Exceeded;

local_DebounceTimer(IN := local_DebounceEnable, PT := DebounceTime);

Weld_Soft_Start_Active := NOT local_PowerUpTimer.Q;
Operator_Alert := Weld_E_Stop_NC AND local_DebounceTimer.Q;

END_FUNCTION_BLOCK

(* ---- public-easy-05.patch_base_02.st ---- *)
FUNCTION_BLOCK WeldGapAlarm
VAR_INPUT
    Gap_Exceeded : BOOL;
    Weld_E_Stop_NC : BOOL;
    DebounceTime : TIME;
END_VAR
VAR_OUTPUT
    Operator_Alert : BOOL;
    Weld_Soft_Start_Active : BOOL;
END_VAR
VAR
    local_PowerUpTimer : TON;
    local_DebounceTimer : TON;
    local_DebounceEnable : BOOL;
END_VAR

(* CONTRACT_RULES [] *)

(* ENGINEERING_CONTRACT
Operator_Alert:
  Activate when E-stop inactive, power-up timer completed, and Gap_Exceeded has been TRUE continuously for DebounceTime.
  Hold while Gap_Exceeded remains TRUE after elapsed DebounceTime.
  Reset immediately on Gap_Exceeded=FALSE, E-stop active, or during initialization.
  Same-scan priority: E-stop active > initialization > debounced gap alarm.
Weld_Soft_Start_Active:
  Activate at power-up and hold TRUE for exactly the 5 s initialization period.
  Deactivate automatically when local_PowerUpTimer reaches 5 s; no manual reset.
  Same-scan priority: independent of E-stop and alarm deactivation.
Units/boundaries: power-up interval = T#5S; DebounceTime is TIME in milliseconds and must be positive.
*)

local_PowerUpTimer(IN := TRUE, PT := T#5S);

local_DebounceEnable := NOT local_PowerUpTimer.Q
                        AND Weld_E_Stop_NC
                        AND Gap_Exceeded;

local_DebounceTimer(IN := local_DebounceEnable, PT := DebounceTime);

Weld_Soft_Start_Active := NOT local_PowerUpTimer.Q;
Operator_Alert := Weld_E_Stop_NC AND local_DebounceTimer.Q;

END_FUNCTION_BLOCK

(* ---- public-easy-05.raw_candidate_01.st ---- *)
FUNCTION_BLOCK WeldGapAlarm
VAR_INPUT
    Gap_Exceeded : BOOL;
    Weld_E_Stop_NC : BOOL;
    DebounceTime : TIME;
END_VAR
VAR_OUTPUT
    Operator_Alert : BOOL;
    Weld_Soft_Start_Active : BOOL;
END_VAR
VAR
    local_PowerUpTimer : TON;
    local_DebounceTimer : TON;
    local_DebounceEnable : BOOL;
END_VAR

(* CONTRACT_RULES [] *)

(* ENGINEERING_CONTRACT
Operator_Alert:
  Activate when E-stop inactive, power-up timer completed, and Gap_Exceeded has been TRUE continuously for DebounceTime.
  Hold while Gap_Exceeded remains TRUE after elapsed DebounceTime.
  Reset immediately on Gap_Exceeded=FALSE, E-stop active, or during initialization.
  Same-scan priority: E-stop active > initialization > debounced gap alarm.
Weld_Soft_Start_Active:
  Activate at power-up and hold TRUE for exactly the 5 s initialization period.
  Deactivate automatically when local_PowerUpTimer reaches 5 s; no manual reset.
  Same-scan priority: independent of E-stop and alarm deactivation.
Units/boundaries: power-up interval = T#5S; DebounceTime is TIME in milliseconds and must be positive.
*)

local_PowerUpTimer(IN := TRUE, PT := T#5S);

local_DebounceEnable := NOT local_PowerUpTimer.Q
                        AND Weld_E_Stop_NC
                        AND Gap_Exceeded;

local_DebounceTimer(IN := local_DebounceEnable, PT := DebounceTime);

Weld_Soft_Start_Active := NOT local_PowerUpTimer.Q;
Operator_Alert := Weld_E_Stop_NC AND local_DebounceTimer.Q;

END_FUNCTION_BLOCK

(* ---- public-easy-05.raw_candidate_02.st ---- *)
FUNCTION_BLOCK WeldGapAlarm
VAR_INPUT
    Gap_Exceeded : BOOL;
    Weld_E_Stop_NC : BOOL;
    DebounceTime : TIME;
END_VAR
VAR_OUTPUT
    Operator_Alert : BOOL;
    Weld_Soft_Start_Active : BOOL;
END_VAR
VAR
    local_PowerUpTimer : TON;
    local_DebounceTimer : TON;
    local_DebounceEnable : BOOL;
END_VAR

(* CONTRACT_RULES [] *)

(* ENGINEERING_CONTRACT
Operator_Alert:
  Activate when E-stop inactive, power-up timer completed, and Gap_Exceeded has been TRUE continuously for DebounceTime.
  Hold while Gap_Exceeded remains TRUE after elapsed DebounceTime.
  Reset immediately on Gap_Exceeded=FALSE, E-stop active, or during initialization.
  Same-scan priority: E-stop active > initialization > debounced gap alarm.
Weld_Soft_Start_Active:
  Activate at power-up and hold TRUE for exactly the 5 s initialization period.
  Deactivate automatically when local_PowerUpTimer reaches 5 s; no manual reset.
  Same-scan priority: independent of E-stop and alarm deactivation.
Units/boundaries: power-up interval = T#5S; DebounceTime is TIME in milliseconds and must be positive.
*)

local_PowerUpTimer(IN := TRUE, PT := T#5S);

local_DebounceEnable := local_PowerUpTimer.Q
                        AND Weld_E_Stop_NC
                        AND Gap_Exceeded;

local_DebounceTimer(IN := local_DebounceEnable, PT := DebounceTime);

Weld_Soft_Start_Active := NOT local_PowerUpTimer.Q;
Operator_Alert := Weld_E_Stop_NC AND local_DebounceTimer.Q;

END_FUNCTION_BLOCK

(* ---- public-easy-06.candidate_01.st ---- *)
FUNCTION_BLOCK AerationBlowerDelayedStart
VAR_INPUT
    DO_LOW : BOOL;
    AERATION_E_STOP_NC : BOOL;
END_VAR
VAR_OUTPUT
    BLOWER_RUN : BOOL := FALSE;
    AERATION_BLOWER_CYCLE_COUNT : UINT := 0;
END_VAR
VAR
    tmp_Demand : BOOL;
    tmp_StartDelay : TON;
    tmp_RunRising : R_TRIG;
END_VAR

(* ENGINEERING_CONTRACT
- Activation: BLOWER_RUN becomes TRUE only after DO_LOW AND AERATION_E_STOP_NC remain TRUE for T#5S [PUB001].
- Retention/hold: BLOWER_RUN remains TRUE while the demand condition stays satisfied; it is not latched [PUB001].
- Reset/deactivation: DO_LOW FALSE or active emergency stop immediately sets BLOWER_RUN FALSE and resets the TON [PUB002].
- Same-scan priority: condition FALSE terminates timing and clears BLOWER_RUN before cycle-edge evaluation [PUB001, PUB002].
- Cycle count: increments once on each FALSE-to-TRUE BLOWER_RUN edge, holds otherwise, and starts at zero [PUB003, PUB004].
- Units/boundaries: 5 seconds, UINT cycle count, BOOL enable only with no speed ramp [PUB001, PUB003, PUB004].
*)

(* CONTRACT_RULES [] *)

tmp_Demand := DO_LOW AND AERATION_E_STOP_NC;

tmp_StartDelay(IN := tmp_Demand, PT := T#5S);
BLOWER_RUN := tmp_StartDelay.Q;

tmp_RunRising(CLK := BLOWER_RUN);
IF tmp_RunRising.Q THEN
    AERATION_BLOWER_CYCLE_COUNT := AERATION_BLOWER_CYCLE_COUNT + 1;
END_IF;

END_FUNCTION_BLOCK

(* ---- public-easy-06.raw_candidate_01.st ---- *)
FUNCTION_BLOCK AerationBlowerDelayedStart
VAR_INPUT
    DO_LOW : BOOL;
    AERATION_E_STOP_NC : BOOL;
END_VAR
VAR_OUTPUT
    BLOWER_RUN : BOOL := FALSE;
    AERATION_BLOWER_CYCLE_COUNT : UINT := 0;
END_VAR
VAR
    tmp_Demand : BOOL;
    tmp_StartDelay : TON;
    tmp_RunRising : R_TRIG;
END_VAR

(* ENGINEERING_CONTRACT
- Activation: BLOWER_RUN becomes TRUE only after DO_LOW AND AERATION_E_STOP_NC remain TRUE for T#5S [PUB001].
- Retention/hold: BLOWER_RUN remains TRUE while the demand condition stays satisfied; it is not latched [PUB001].
- Reset/deactivation: DO_LOW FALSE or active emergency stop immediately sets BLOWER_RUN FALSE and resets the TON [PUB002].
- Same-scan priority: condition FALSE terminates timing and clears BLOWER_RUN before cycle-edge evaluation [PUB001, PUB002].
- Cycle count: increments once on each FALSE-to-TRUE BLOWER_RUN edge, holds otherwise, and starts at zero [PUB003, PUB004].
- Units/boundaries: 5 seconds, UINT cycle count, BOOL enable only with no speed ramp [PUB001, PUB003, PUB004].
*)

(* CONTRACT_RULES [] *)

tmp_Demand := DO_LOW AND AERATION_E_STOP_NC;

tmp_StartDelay(IN := tmp_Demand, PT := T#5S);
BLOWER_RUN := tmp_StartDelay.Q;

tmp_RunRising(CLK := BLOWER_RUN);
IF tmp_RunRising.Q THEN
    AERATION_BLOWER_CYCLE_COUNT := AERATION_BLOWER_CYCLE_COUNT + 1;
END_IF;

END_FUNCTION_BLOCK

(* ---- public-hard-01.candidate_01.st ---- *)
(* CONTRACT_RULES [] *)

(* ENGINEERING_CONTRACT
   - ESTOP: ESTOP=FALSE forces every output OFF in this scan; manual and auto commands are inhibited.
   - Manual runs: only while OpeMode=FALSE and ESTOP=TRUE; each start button rising edge toggles its retained output latch.
   - Auto sequence: AUTOSTART rising edge while OpeMode=TRUE enters FILL_A; output valves follow the sequence below.
   - Valve A: ON in FILL_A; Level>=50 closes A and opens B (PUB012).
   - Valve B: ON in FILL_B; Level>=80 closes B (PUB012/PUB013).
   - ProcessMode=FALSE: at Level>=80 mixer starts; MixMotorComplete latches completion, then mixer off and Valve D ON, sequence done (PUB014).
   - ProcessMode=TRUE: at Level>=80 Valve C opens; Level>=100 closes C and starts mixer; completion opens D (PUB014).
   - Mix complete is latched until the next AUTOSTART; Valve D remains ON in DONE because no stop/reset is stated.
   - Thresholds are inclusive >=; Level is INT cm; PROCESSMODE is read live at the 80 cm transition.
*)

TYPE E_MaterialProportioningState :
(
    MP_IDLE,
    MP_FILL_A,
    MP_FILL_B,
    MP_MIX_SIMPLE,
    MP_FILL_C,
    MP_MIX_C,
    MP_DONE
) := MP_IDLE;
END_TYPE;

FUNCTION_BLOCK MaterialProportioningControl
VAR_INPUT
    estop : BOOL;
    opeMode : BOOL;
    valveAStart : BOOL;
    valveBStart : BOOL;
    valveCStart : BOOL;
    valveDStart : BOOL;
    mixMotorStart : BOOL;
    autoStart : BOOL;
    processMode : BOOL;
    levelSensor : INT;
    mixMotorComplete : BOOL;
END_VAR
VAR_OUTPUT
    valveARun : BOOL;
    valveBRun : BOOL;
    valveCRun : BOOL;
    valveDRun : BOOL;
    mixMotorRun : BOOL;
END_VAR
VAR
    tmp_trigValveA : R_TRIG;
    tmp_trigValveB : R_TRIG;
    tmp_trigValveC : R_TRIG;
    tmp_trigValveD : R_TRIG;
    tmp_trigMixMotor : R_TRIG;
    tmp_trigAutoStart : R_TRIG;

    manualValveARun : BOOL := FALSE;
    manualValveBRun : BOOL := FALSE;
    manualValveCRun : BOOL := FALSE;
    manualValveDRun : BOOL := FALSE;
    manualMixMotorRun : BOOL := FALSE;

    state : E_MaterialProportioningState := MP_IDLE;
    mixCompleteLatched : BOOL := FALSE;
END_VAR

tmp_trigValveA(CLK := valveAStart);
tmp_trigValveB(CLK := valveBStart);
tmp_trigValveC(CLK := valveCStart);
tmp_trigValveD(CLK := valveDStart);
tmp_trigMixMotor(CLK := mixMotorStart);
tmp_trigAutoStart(CLK := autoStart);

IF NOT estop THEN
    valveARun := FALSE;
    valveBRun := FALSE;
    valveCRun := FALSE;
    valveDRun := FALSE;
    mixMotorRun := FALSE;

ELSIF NOT opeMode THEN
    state := MP_IDLE;
    mixCompleteLatched := FALSE;

    IF tmp_trigValveA.Q THEN
        manualValveARun := NOT manualValveARun;
    END_IF;
    IF tmp_trigValveB.Q THEN
        manualValveBRun := NOT manualValveBRun;
    END_IF;
    IF tmp_trigValveC.Q THEN
        manualValveCRun := NOT manualValveCRun;
    END_IF;
    IF tmp_trigValveD.Q THEN
        manualValveDRun := NOT manualValveDRun;
    END_IF;
    IF tmp_trigMixMotor.Q THEN
        manualMixMotorRun := NOT manualMixMotorRun;
    END_IF;

    valveARun := manualValveARun;
    valveBRun := manualValveBRun;
    valveCRun := manualValveCRun;
    valveDRun := manualValveDRun;
    mixMotorRun := manualMixMotorRun;

ELSE
    IF tmp_trigAutoStart.Q THEN
        state := MP_FILL_A;
        mixCompleteLatched := FALSE;
    END_IF;

    CASE state OF
        MP_IDLE:
            valveARun := FALSE;
            valveBRun := FALSE;
            valveCRun := FALSE;
            valveDRun := FALSE;
            mixMotorRun := FALSE;

        MP_FILL_A:
            valveARun := TRUE;
            valveBRun := FALSE;
            valveCRun := FALSE;
            valveDRun := FALSE;
            mixMotorRun := FALSE;

            IF levelSensor >= 50 THEN
                valveARun := FALSE;
                valveBRun := TRUE;
                state := MP_FILL_B;
            END_IF;

        MP_FILL_B:
            valveARun := FALSE;
            valveBRun := TRUE;
            valveCRun := FALSE;
            valveDRun := FALSE;
            mixMotorRun := FALSE;

            IF levelSensor >= 80 THEN
                valveBRun := FALSE;
                IF NOT processMode THEN
                    mixMotorRun := TRUE;
                    mixCompleteLatched := FALSE;
                    state := MP_MIX_SIMPLE;
                ELSE
                    valveCRun := TRUE;
                    state := MP_FILL_C;
                END_IF;
            END_IF;

        MP_FILL_C:
            valveARun := FALSE;
            valveBRun := FALSE;
            valveCRun := TRUE;
            valveDRun := FALSE;
            mixMotorRun := FALSE;

            IF levelSensor >= 100 THEN
                valveCRun := FALSE;
                mixMotorRun := TRUE;
                mixCompleteLatched := FALSE;
                state := MP_MIX_C;
            END_IF;

        MP_MIX_SIMPLE:
            valveARun := FALSE;
            valveBRun := FALSE;
            valveCRun := FALSE;
            valveDRun := FALSE;
            mixMotorRun := TRUE;

            IF mixMotorComplete THEN
                mixCompleteLatched := TRUE;
            END_IF;

            IF mixCompleteLatched THEN
                mixMotorRun := FALSE;
                valveDRun := TRUE;
                state := MP_DONE;
            END_IF;

        MP_MIX_C:
            valveARun := FALSE;
            valveBRun := FALSE;
            valveCRun := FALSE;
            valveDRun := FALSE;
            mixMotorRun := TRUE;

            IF mixMotorComplete THEN
                mixCompleteLatched := TRUE;
            END_IF;

            IF mixCompleteLatched THEN
                mixMotorRun := FALSE;
                valveDRun := TRUE;
                state := MP_DONE;
            END_IF;

        MP_DONE:
            valveARun := FALSE;
            valveBRun := FALSE;
            valveCRun := FALSE;
            valveDRun := TRUE;
            mixMotorRun := FALSE;
    END_CASE;
END_IF;
END_FUNCTION_BLOCK

(* ---- public-hard-01.candidate_02.st ---- *)
(* CONTRACT_RULES [] *)

(* ENGINEERING_CONTRACT
   - ESTOP: ESTOP=FALSE forces every output OFF in this scan; manual and auto commands are inhibited.
   - Manual runs: only while OpeMode=FALSE and ESTOP=TRUE; each start button rising edge toggles its retained output latch.
   - Auto sequence: AUTOSTART rising edge while OpeMode=TRUE enters FILL_A; output valves follow the sequence below.
   - Valve A: ON in FILL_A; Level>=50 closes A and opens B (PUB012).
   - Valve B: ON in FILL_B; Level>=80 closes B (PUB012/PUB013).
   - ProcessMode=FALSE: at Level>=80 mixer starts; MixMotorComplete latches completion, then mixer off and Valve D ON, sequence done (PUB014).
   - ProcessMode=TRUE: at Level>=80 Valve C opens; Level>=100 closes C and starts mixer; completion opens D (PUB014).
   - Mix complete is latched until the next AUTOSTART; Valve D remains ON in DONE because no stop/reset is stated.
   - Thresholds are inclusive >=; Level is INT cm; PROCESSMODE is read live at the 80 cm transition.
*)

TYPE E_MaterialProportioningState :
(
    MP_IDLE,
    MP_FILL_A,
    MP_FILL_B,
    MP_MIX_SIMPLE,
    MP_FILL_C,
    MP_MIX_C,
    MP_DONE
) := MP_IDLE;
END_TYPE;

FUNCTION_BLOCK MaterialProportioningControl
VAR_INPUT
    estop : BOOL;
    opeMode : BOOL;
    valveAStart : BOOL;
    valveBStart : BOOL;
    valveCStart : BOOL;
    valveDStart : BOOL;
    mixMotorStart : BOOL;
    autoStart : BOOL;
    processMode : BOOL;
    levelSensor : INT;
    mixMotorComplete : BOOL;
END_VAR
VAR_OUTPUT
    valveARun : BOOL;
    valveBRun : BOOL;
    valveCRun : BOOL;
    valveDRun : BOOL;
    mixMotorRun : BOOL;
END_VAR
VAR
    tmp_trigValveA : R_TRIG;
    tmp_trigValveB : R_TRIG;
    tmp_trigValveC : R_TRIG;
    tmp_trigValveD : R_TRIG;
    tmp_trigMixMotor : R_TRIG;
    tmp_trigAutoStart : R_TRIG;

    manualValveARun : BOOL := FALSE;
    manualValveBRun : BOOL := FALSE;
    manualValveCRun : BOOL := FALSE;
    manualValveDRun : BOOL := FALSE;
    manualMixMotorRun : BOOL := FALSE;

    state : E_MaterialProportioningState := MP_IDLE;
    mixCompleteLatched : BOOL := FALSE;
END_VAR

tmp_trigValveA(CLK := valveAStart);
tmp_trigValveB(CLK := valveBStart);
tmp_trigValveC(CLK := valveCStart);
tmp_trigValveD(CLK := valveDStart);
tmp_trigMixMotor(CLK := mixMotorStart);
tmp_trigAutoStart(CLK := autoStart);

IF NOT estop THEN
    valveARun := FALSE;
    valveBRun := FALSE;
    valveCRun := FALSE;
    valveDRun := FALSE;
    mixMotorRun := FALSE;

ELSIF NOT opeMode THEN
    state := MP_IDLE;
    mixCompleteLatched := FALSE;

    IF tmp_trigValveA.Q THEN
        manualValveARun := NOT manualValveARun;
    END_IF;
    IF tmp_trigValveB.Q THEN
        manualValveBRun := NOT manualValveBRun;
    END_IF;
    IF tmp_trigValveC.Q THEN
        manualValveCRun := NOT manualValveCRun;
    END_IF;
    IF tmp_trigValveD.Q THEN
        manualValveDRun := NOT manualValveDRun;
    END_IF;
    IF tmp_trigMixMotor.Q THEN
        manualMixMotorRun := NOT manualMixMotorRun;
    END_IF;

    valveARun := manualValveARun;
    valveBRun := manualValveBRun;
    valveCRun := manualValveCRun;
    valveDRun := manualValveDRun;
    mixMotorRun := manualMixMotorRun;

ELSE
    IF tmp_trigAutoStart.Q THEN
        state := MP_FILL_A;
        mixCompleteLatched := FALSE;
    END_IF;

    CASE state OF
        MP_IDLE:
            valveARun := FALSE;
            valveBRun := FALSE;
            valveCRun := FALSE;
            valveDRun := FALSE;
            mixMotorRun := FALSE;

        MP_FILL_A:
            valveARun := TRUE;
            valveBRun := FALSE;
            valveCRun := FALSE;
            valveDRun := FALSE;
            mixMotorRun := FALSE;

            IF levelSensor >= 50 THEN
                valveARun := FALSE;
                valveBRun := TRUE;
                state := MP_FILL_B;
            END_IF;

        MP_FILL_B:
            valveARun := FALSE;
            valveBRun := TRUE;
            valveCRun := FALSE;
            valveDRun := FALSE;
            mixMotorRun := FALSE;

            IF levelSensor >= 80 THEN
                valveBRun := FALSE;
                IF NOT processMode THEN
                    mixMotorRun := TRUE;
                    mixCompleteLatched := FALSE;
                    state := MP_MIX_SIMPLE;
                ELSE
                    IF levelSensor >= 100 THEN
                        valveCRun := FALSE;
                        mixMotorRun := TRUE;
                        mixCompleteLatched := FALSE;
                        state := MP_MIX_C;
                    ELSE
                        valveCRun := TRUE;
                        state := MP_FILL_C;
                    END_IF;
                END_IF;
            END_IF;

        MP_FILL_C:
            valveARun := FALSE;
            valveBRun := FALSE;
            valveCRun := TRUE;
            valveDRun := FALSE;
            mixMotorRun := FALSE;

            IF levelSensor >= 100 THEN
                valveCRun := FALSE;
                mixMotorRun := TRUE;
                mixCompleteLatched := FALSE;
                state := MP_MIX_C;
            END_IF;

        MP_MIX_SIMPLE:
            valveARun := FALSE;
            valveBRun := FALSE;
            valveCRun := FALSE;
            valveDRun := FALSE;
            mixMotorRun := TRUE;

            IF mixMotorComplete THEN
                mixCompleteLatched := TRUE;
            END_IF;

            IF mixCompleteLatched THEN
                mixMotorRun := FALSE;
                valveDRun := TRUE;
                state := MP_DONE;
            END_IF;

        MP_MIX_C:
            valveARun := FALSE;
            valveBRun := FALSE;
            valveCRun := FALSE;
            valveDRun := FALSE;
            mixMotorRun := TRUE;

            IF mixMotorComplete THEN
                mixCompleteLatched := TRUE;
            END_IF;

            IF mixCompleteLatched THEN
                mixMotorRun := FALSE;
                valveDRun := TRUE;
                state := MP_DONE;
            END_IF;

        MP_DONE:
            valveARun := FALSE;
            valveBRun := FALSE;
            valveCRun := FALSE;
            valveDRun := TRUE;
            mixMotorRun := FALSE;
    END_CASE;
END_IF;
END_FUNCTION_BLOCK

(* ---- public-hard-01.candidate_03.st ---- *)
(* CONTRACT_RULES [] *)

(* ENGINEERING_CONTRACT
   - ESTOP: ESTOP=FALSE forces every output OFF in this scan; manual and auto commands are inhibited.
   - Manual runs: only while OpeMode=FALSE and ESTOP=TRUE; each start button rising edge toggles its retained output latch.
   - Auto sequence: AUTOSTART rising edge while OpeMode=TRUE enters FILL_A; output valves follow the sequence below.
   - Valve A: ON in FILL_A; Level>=50 closes A and opens B (PUB012).
   - Valve B: ON in FILL_B; Level>=80 closes B (PUB012/PUB013).
   - ProcessMode=FALSE: at Level>=80 mixer starts; MixMotorComplete latches completion, then mixer off and Valve D ON, sequence done (PUB014).
   - ProcessMode=TRUE: at Level>=80 Valve C opens; Level>=100 closes C and starts mixer; completion opens D (PUB014).
   - Mix complete is latched until the next AUTOSTART; Valve D remains ON in DONE because no stop/reset is stated.
   - Thresholds are inclusive >=; Level is INT cm; PROCESSMODE is read live at the 80 cm transition.
*)

TYPE E_MaterialProportioningState :
(
    MP_IDLE,
    MP_FILL_A,
    MP_FILL_B,
    MP_MIX_SIMPLE,
    MP_FILL_C,
    MP_MIX_C,
    MP_DONE
) := MP_IDLE;
END_TYPE;

FUNCTION_BLOCK MaterialProportioningControl
VAR_INPUT
    estop : BOOL;
    opeMode : BOOL;
    valveAStart : BOOL;
    valveBStart : BOOL;
    valveCStart : BOOL;
    valveDStart : BOOL;
    mixMotorStart : BOOL;
    autoStart : BOOL;
    processMode : BOOL;
    levelSensor : INT;
    mixMotorComplete : BOOL;
END_VAR
VAR_OUTPUT
    valveARun : BOOL;
    valveBRun : BOOL;
    valveCRun : BOOL;
    valveDRun : BOOL;
    mixMotorRun : BOOL;
END_VAR
VAR
    tmp_trigValveA : R_TRIG;
    tmp_trigValveB : R_TRIG;
    tmp_trigValveC : R_TRIG;
    tmp_trigValveD : R_TRIG;
    tmp_trigMixMotor : R_TRIG;
    tmp_trigAutoStart : R_TRIG;

    manualValveARun : BOOL := FALSE;
    manualValveBRun : BOOL := FALSE;
    manualValveCRun : BOOL := FALSE;
    manualValveDRun : BOOL := FALSE;
    manualMixMotorRun : BOOL := FALSE;

    state : E_MaterialProportioningState := MP_IDLE;
    mixCompleteLatched : BOOL := FALSE;
END_VAR

tmp_trigValveA(CLK := valveAStart);
tmp_trigValveB(CLK := valveBStart);
tmp_trigValveC(CLK := valveCStart);
tmp_trigValveD(CLK := valveDStart);
tmp_trigMixMotor(CLK := mixMotorStart);
tmp_trigAutoStart(CLK := autoStart);

IF NOT estop THEN
    valveARun := FALSE;
    valveBRun := FALSE;
    valveCRun := FALSE;
    valveDRun := FALSE;
    mixMotorRun := FALSE;

ELSIF NOT opeMode THEN
    state := MP_IDLE;
    mixCompleteLatched := FALSE;

    IF tmp_trigValveA.Q THEN
        manualValveARun := NOT manualValveARun;
    END_IF;
    IF tmp_trigValveB.Q THEN
        manualValveBRun := NOT manualValveBRun;
    END_IF;
    IF tmp_trigValveC.Q THEN
        manualValveCRun := NOT manualValveCRun;
    END_IF;
    IF tmp_trigValveD.Q THEN
        manualValveDRun := NOT manualValveDRun;
    END_IF;
    IF tmp_trigMixMotor.Q THEN
        manualMixMotorRun := NOT manualMixMotorRun;
    END_IF;

    valveARun := manualValveARun;
    valveBRun := manualValveBRun;
    valveCRun := manualValveCRun;
    valveDRun := manualValveDRun;
    mixMotorRun := manualMixMotorRun;

ELSE
    IF tmp_trigAutoStart.Q THEN
        state := MP_FILL_A;
        mixCompleteLatched := FALSE;
    END_IF;

    CASE state OF
        MP_IDLE:
            valveARun := FALSE;
            valveBRun := FALSE;
            valveCRun := FALSE;
            valveDRun := FALSE;
            mixMotorRun := FALSE;

        MP_FILL_A:
            valveARun := TRUE;
            valveBRun := FALSE;
            valveCRun := FALSE;
            valveDRun := FALSE;
            mixMotorRun := FALSE;

            IF levelSensor >= 80 THEN
                valveARun := FALSE;
                valveBRun := FALSE;
                IF NOT processMode THEN
                    mixMotorRun := TRUE;
                    mixCompleteLatched := FALSE;
                    state := MP_MIX_SIMPLE;
                ELSIF levelSensor >= 100 THEN
                    valveCRun := FALSE;
                    mixMotorRun := TRUE;
                    mixCompleteLatched := FALSE;
                    state := MP_MIX_C;
                ELSE
                    valveCRun := TRUE;
                    state := MP_FILL_C;
                END_IF;
            ELSIF levelSensor >= 50 THEN
                valveARun := FALSE;
                valveBRun := TRUE;
                state := MP_FILL_B;
            END_IF;

        MP_FILL_B:
            valveARun := FALSE;
            valveBRun := TRUE;
            valveCRun := FALSE;
            valveDRun := FALSE;
            mixMotorRun := FALSE;

            IF levelSensor >= 80 THEN
                valveBRun := FALSE;
                IF NOT processMode THEN
                    mixMotorRun := TRUE;
                    mixCompleteLatched := FALSE;
                    state := MP_MIX_SIMPLE;
                ELSE
                    IF levelSensor >= 100 THEN
                        valveCRun := FALSE;
                        mixMotorRun := TRUE;
                        mixCompleteLatched := FALSE;
                        state := MP_MIX_C;
                    ELSE
                        valveCRun := TRUE;
                        state := MP_FILL_C;
                    END_IF;
                END_IF;
            END_IF;

        MP_FILL_C:
            valveARun := FALSE;
            valveBRun := FALSE;
            valveCRun := TRUE;
            valveDRun := FALSE;
            mixMotorRun := FALSE;

            IF levelSensor >= 100 THEN
                valveCRun := FALSE;
                mixMotorRun := TRUE;
                mixCompleteLatched := FALSE;
                state := MP_MIX_C;
            END_IF;

        MP_MIX_SIMPLE:
            valveARun := FALSE;
            valveBRun := FALSE;
            valveCRun := FALSE;
            valveDRun := FALSE;
            mixMotorRun := TRUE;

            IF mixMotorComplete THEN
                mixCompleteLatched := TRUE;
            END_IF;

            IF mixCompleteLatched THEN
                mixMotorRun := FALSE;
                valveDRun := TRUE;
                state := MP_DONE;
            END_IF;

        MP_MIX_C:
            valveARun := FALSE;
            valveBRun := FALSE;
            valveCRun := FALSE;
            valveDRun := FALSE;
            mixMotorRun := TRUE;

            IF mixMotorComplete THEN
                mixCompleteLatched := TRUE;
            END_IF;

            IF mixCompleteLatched THEN
                mixMotorRun := FALSE;
                valveDRun := TRUE;
                state := MP_DONE;
            END_IF;

        MP_DONE:
            valveARun := FALSE;
            valveBRun := FALSE;
            valveCRun := FALSE;
            valveDRun := TRUE;
            mixMotorRun := FALSE;
    END_CASE;
END_IF;
END_FUNCTION_BLOCK

(* ---- public-hard-01.patch_base_02.st ---- *)
(* CONTRACT_RULES [] *)

(* ENGINEERING_CONTRACT
   - ESTOP: ESTOP=FALSE forces every output OFF in this scan; manual and auto commands are inhibited.
   - Manual runs: only while OpeMode=FALSE and ESTOP=TRUE; each start button rising edge toggles its retained output latch.
   - Auto sequence: AUTOSTART rising edge while OpeMode=TRUE enters FILL_A; output valves follow the sequence below.
   - Valve A: ON in FILL_A; Level>=50 closes A and opens B (PUB012).
   - Valve B: ON in FILL_B; Level>=80 closes B (PUB012/PUB013).
   - ProcessMode=FALSE: at Level>=80 mixer starts; MixMotorComplete latches completion, then mixer off and Valve D ON, sequence done (PUB014).
   - ProcessMode=TRUE: at Level>=80 Valve C opens; Level>=100 closes C and starts mixer; completion opens D (PUB014).
   - Mix complete is latched until the next AUTOSTART; Valve D remains ON in DONE because no stop/reset is stated.
   - Thresholds are inclusive >=; Level is INT cm; PROCESSMODE is read live at the 80 cm transition.
*)

TYPE E_MaterialProportioningState :
(
    MP_IDLE,
    MP_FILL_A,
    MP_FILL_B,
    MP_MIX_SIMPLE,
    MP_FILL_C,
    MP_MIX_C,
    MP_DONE
) := MP_IDLE;
END_TYPE;

FUNCTION_BLOCK MaterialProportioningControl
VAR_INPUT
    estop : BOOL;
    opeMode : BOOL;
    valveAStart : BOOL;
    valveBStart : BOOL;
    valveCStart : BOOL;
    valveDStart : BOOL;
    mixMotorStart : BOOL;
    autoStart : BOOL;
    processMode : BOOL;
    levelSensor : INT;
    mixMotorComplete : BOOL;
END_VAR
VAR_OUTPUT
    valveARun : BOOL;
    valveBRun : BOOL;
    valveCRun : BOOL;
    valveDRun : BOOL;
    mixMotorRun : BOOL;
END_VAR
VAR
    tmp_trigValveA : R_TRIG;
    tmp_trigValveB : R_TRIG;
    tmp_trigValveC : R_TRIG;
    tmp_trigValveD : R_TRIG;
    tmp_trigMixMotor : R_TRIG;
    tmp_trigAutoStart : R_TRIG;

    manualValveARun : BOOL := FALSE;
    manualValveBRun : BOOL := FALSE;
    manualValveCRun : BOOL := FALSE;
    manualValveDRun : BOOL := FALSE;
    manualMixMotorRun : BOOL := FALSE;

    state : E_MaterialProportioningState := MP_IDLE;
    mixCompleteLatched : BOOL := FALSE;
END_VAR

tmp_trigValveA(CLK := valveAStart);
tmp_trigValveB(CLK := valveBStart);
tmp_trigValveC(CLK := valveCStart);
tmp_trigValveD(CLK := valveDStart);
tmp_trigMixMotor(CLK := mixMotorStart);
tmp_trigAutoStart(CLK := autoStart);

IF NOT estop THEN
    valveARun := FALSE;
    valveBRun := FALSE;
    valveCRun := FALSE;
    valveDRun := FALSE;
    mixMotorRun := FALSE;

ELSIF NOT opeMode THEN
    state := MP_IDLE;
    mixCompleteLatched := FALSE;

    IF tmp_trigValveA.Q THEN
        manualValveARun := NOT manualValveARun;
    END_IF;
    IF tmp_trigValveB.Q THEN
        manualValveBRun := NOT manualValveBRun;
    END_IF;
    IF tmp_trigValveC.Q THEN
        manualValveCRun := NOT manualValveCRun;
    END_IF;
    IF tmp_trigValveD.Q THEN
        manualValveDRun := NOT manualValveDRun;
    END_IF;
    IF tmp_trigMixMotor.Q THEN
        manualMixMotorRun := NOT manualMixMotorRun;
    END_IF;

    valveARun := manualValveARun;
    valveBRun := manualValveBRun;
    valveCRun := manualValveCRun;
    valveDRun := manualValveDRun;
    mixMotorRun := manualMixMotorRun;

ELSE
    IF tmp_trigAutoStart.Q THEN
        state := MP_FILL_A;
        mixCompleteLatched := FALSE;
    END_IF;

    CASE state OF
        MP_IDLE:
            valveARun := FALSE;
            valveBRun := FALSE;
            valveCRun := FALSE;
            valveDRun := FALSE;
            mixMotorRun := FALSE;

        MP_FILL_A:
            valveARun := TRUE;
            valveBRun := FALSE;
            valveCRun := FALSE;
            valveDRun := FALSE;
            mixMotorRun := FALSE;

            IF levelSensor >= 50 THEN
                valveARun := FALSE;
                valveBRun := TRUE;
                state := MP_FILL_B;
            END_IF;

        MP_FILL_B:
            valveARun := FALSE;
            valveBRun := TRUE;
            valveCRun := FALSE;
            valveDRun := FALSE;
            mixMotorRun := FALSE;

            IF levelSensor >= 80 THEN
                valveBRun := FALSE;
                IF NOT processMode THEN
                    mixMotorRun := TRUE;
                    mixCompleteLatched := FALSE;
                    state := MP_MIX_SIMPLE;
                ELSE
                    valveCRun := TRUE;
                    state := MP_FILL_C;
                END_IF;
            END_IF;

        MP_FILL_C:
            valveARun := FALSE;
            valveBRun := FALSE;
            valveCRun := TRUE;
            valveDRun := FALSE;
            mixMotorRun := FALSE;

            IF levelSensor >= 100 THEN
                valveCRun := FALSE;
                mixMotorRun := TRUE;
                mixCompleteLatched := FALSE;
                state := MP_MIX_C;
            END_IF;

        MP_MIX_SIMPLE:
            valveARun := FALSE;
            valveBRun := FALSE;
            valveCRun := FALSE;
            valveDRun := FALSE;
            mixMotorRun := TRUE;

            IF mixMotorComplete THEN
                mixCompleteLatched := TRUE;
            END_IF;

            IF mixCompleteLatched THEN
                mixMotorRun := FALSE;
                valveDRun := TRUE;
                state := MP_DONE;
            END_IF;

        MP_MIX_C:
            valveARun := FALSE;
            valveBRun := FALSE;
            valveCRun := FALSE;
            valveDRun := FALSE;
            mixMotorRun := TRUE;

            IF mixMotorComplete THEN
                mixCompleteLatched := TRUE;
            END_IF;

            IF mixCompleteLatched THEN
                mixMotorRun := FALSE;
                valveDRun := TRUE;
                state := MP_DONE;
            END_IF;

        MP_DONE:
            valveARun := FALSE;
            valveBRun := FALSE;
            valveCRun := FALSE;
            valveDRun := TRUE;
            mixMotorRun := FALSE;
    END_CASE;
END_IF;
END_FUNCTION_BLOCK

(* ---- public-hard-01.patch_base_03.st ---- *)
(* CONTRACT_RULES [] *)

(* ENGINEERING_CONTRACT
   - ESTOP: ESTOP=FALSE forces every output OFF in this scan; manual and auto commands are inhibited.
   - Manual runs: only while OpeMode=FALSE and ESTOP=TRUE; each start button rising edge toggles its retained output latch.
   - Auto sequence: AUTOSTART rising edge while OpeMode=TRUE enters FILL_A; output valves follow the sequence below.
   - Valve A: ON in FILL_A; Level>=50 closes A and opens B (PUB012).
   - Valve B: ON in FILL_B; Level>=80 closes B (PUB012/PUB013).
   - ProcessMode=FALSE: at Level>=80 mixer starts; MixMotorComplete latches completion, then mixer off and Valve D ON, sequence done (PUB014).
   - ProcessMode=TRUE: at Level>=80 Valve C opens; Level>=100 closes C and starts mixer; completion opens D (PUB014).
   - Mix complete is latched until the next AUTOSTART; Valve D remains ON in DONE because no stop/reset is stated.
   - Thresholds are inclusive >=; Level is INT cm; PROCESSMODE is read live at the 80 cm transition.
*)

TYPE E_MaterialProportioningState :
(
    MP_IDLE,
    MP_FILL_A,
    MP_FILL_B,
    MP_MIX_SIMPLE,
    MP_FILL_C,
    MP_MIX_C,
    MP_DONE
) := MP_IDLE;
END_TYPE;

FUNCTION_BLOCK MaterialProportioningControl
VAR_INPUT
    estop : BOOL;
    opeMode : BOOL;
    valveAStart : BOOL;
    valveBStart : BOOL;
    valveCStart : BOOL;
    valveDStart : BOOL;
    mixMotorStart : BOOL;
    autoStart : BOOL;
    processMode : BOOL;
    levelSensor : INT;
    mixMotorComplete : BOOL;
END_VAR
VAR_OUTPUT
    valveARun : BOOL;
    valveBRun : BOOL;
    valveCRun : BOOL;
    valveDRun : BOOL;
    mixMotorRun : BOOL;
END_VAR
VAR
    tmp_trigValveA : R_TRIG;
    tmp_trigValveB : R_TRIG;
    tmp_trigValveC : R_TRIG;
    tmp_trigValveD : R_TRIG;
    tmp_trigMixMotor : R_TRIG;
    tmp_trigAutoStart : R_TRIG;

    manualValveARun : BOOL := FALSE;
    manualValveBRun : BOOL := FALSE;
    manualValveCRun : BOOL := FALSE;
    manualValveDRun : BOOL := FALSE;
    manualMixMotorRun : BOOL := FALSE;

    state : E_MaterialProportioningState := MP_IDLE;
    mixCompleteLatched : BOOL := FALSE;
END_VAR

tmp_trigValveA(CLK := valveAStart);
tmp_trigValveB(CLK := valveBStart);
tmp_trigValveC(CLK := valveCStart);
tmp_trigValveD(CLK := valveDStart);
tmp_trigMixMotor(CLK := mixMotorStart);
tmp_trigAutoStart(CLK := autoStart);

IF NOT estop THEN
    valveARun := FALSE;
    valveBRun := FALSE;
    valveCRun := FALSE;
    valveDRun := FALSE;
    mixMotorRun := FALSE;

ELSIF NOT opeMode THEN
    state := MP_IDLE;
    mixCompleteLatched := FALSE;

    IF tmp_trigValveA.Q THEN
        manualValveARun := NOT manualValveARun;
    END_IF;
    IF tmp_trigValveB.Q THEN
        manualValveBRun := NOT manualValveBRun;
    END_IF;
    IF tmp_trigValveC.Q THEN
        manualValveCRun := NOT manualValveCRun;
    END_IF;
    IF tmp_trigValveD.Q THEN
        manualValveDRun := NOT manualValveDRun;
    END_IF;
    IF tmp_trigMixMotor.Q THEN
        manualMixMotorRun := NOT manualMixMotorRun;
    END_IF;

    valveARun := manualValveARun;
    valveBRun := manualValveBRun;
    valveCRun := manualValveCRun;
    valveDRun := manualValveDRun;
    mixMotorRun := manualMixMotorRun;

ELSE
    IF tmp_trigAutoStart.Q THEN
        state := MP_FILL_A;
        mixCompleteLatched := FALSE;
    END_IF;

    CASE state OF
        MP_IDLE:
            valveARun := FALSE;
            valveBRun := FALSE;
            valveCRun := FALSE;
            valveDRun := FALSE;
            mixMotorRun := FALSE;

        MP_FILL_A:
            valveARun := TRUE;
            valveBRun := FALSE;
            valveCRun := FALSE;
            valveDRun := FALSE;
            mixMotorRun := FALSE;

            IF levelSensor >= 50 THEN
                valveARun := FALSE;
                valveBRun := TRUE;
                state := MP_FILL_B;
            END_IF;

        MP_FILL_B:
            valveARun := FALSE;
            valveBRun := TRUE;
            valveCRun := FALSE;
            valveDRun := FALSE;
            mixMotorRun := FALSE;

            IF levelSensor >= 80 THEN
                valveBRun := FALSE;
                IF NOT processMode THEN
                    mixMotorRun := TRUE;
                    mixCompleteLatched := FALSE;
                    state := MP_MIX_SIMPLE;
                ELSE
                    IF levelSensor >= 100 THEN
                        valveCRun := FALSE;
                        mixMotorRun := TRUE;
                        mixCompleteLatched := FALSE;
                        state := MP_MIX_C;
                    ELSE
                        valveCRun := TRUE;
                        state := MP_FILL_C;
                    END_IF;
                END_IF;
            END_IF;

        MP_FILL_C:
            valveARun := FALSE;
            valveBRun := FALSE;
            valveCRun := TRUE;
            valveDRun := FALSE;
            mixMotorRun := FALSE;

            IF levelSensor >= 100 THEN
                valveCRun := FALSE;
                mixMotorRun := TRUE;
                mixCompleteLatched := FALSE;
                state := MP_MIX_C;
            END_IF;

        MP_MIX_SIMPLE:
            valveARun := FALSE;
            valveBRun := FALSE;
            valveCRun := FALSE;
            valveDRun := FALSE;
            mixMotorRun := TRUE;

            IF mixMotorComplete THEN
                mixCompleteLatched := TRUE;
            END_IF;

            IF mixCompleteLatched THEN
                mixMotorRun := FALSE;
                valveDRun := TRUE;
                state := MP_DONE;
            END_IF;

        MP_MIX_C:
            valveARun := FALSE;
            valveBRun := FALSE;
            valveCRun := FALSE;
            valveDRun := FALSE;
            mixMotorRun := TRUE;

            IF mixMotorComplete THEN
                mixCompleteLatched := TRUE;
            END_IF;

            IF mixCompleteLatched THEN
                mixMotorRun := FALSE;
                valveDRun := TRUE;
                state := MP_DONE;
            END_IF;

        MP_DONE:
            valveARun := FALSE;
            valveBRun := FALSE;
            valveCRun := FALSE;
            valveDRun := TRUE;
            mixMotorRun := FALSE;
    END_CASE;
END_IF;
END_FUNCTION_BLOCK

(* ---- public-hard-01.raw_candidate_01.st ---- *)
(* CONTRACT_RULES [] *)

(* ENGINEERING_CONTRACT
   - ESTOP: ESTOP=FALSE forces every output OFF in this scan; manual and auto commands are inhibited.
   - Manual runs: only while OpeMode=FALSE and ESTOP=TRUE; each start button rising edge toggles its retained output latch.
   - Auto sequence: AUTOSTART rising edge while OpeMode=TRUE enters FILL_A; output valves follow the sequence below.
   - Valve A: ON in FILL_A; Level>=50 closes A and opens B (PUB012).
   - Valve B: ON in FILL_B; Level>=80 closes B (PUB012/PUB013).
   - ProcessMode=FALSE: at Level>=80 mixer starts; MixMotorComplete latches completion, then mixer off and Valve D ON, sequence done (PUB014).
   - ProcessMode=TRUE: at Level>=80 Valve C opens; Level>=100 closes C and starts mixer; completion opens D (PUB014).
   - Mix complete is latched until the next AUTOSTART; Valve D remains ON in DONE because no stop/reset is stated.
   - Thresholds are inclusive >=; Level is INT cm; PROCESSMODE is read live at the 80 cm transition.
*)

TYPE E_MaterialProportioningState :
(
    MP_IDLE,
    MP_FILL_A,
    MP_FILL_B,
    MP_MIX_SIMPLE,
    MP_FILL_C,
    MP_MIX_C,
    MP_DONE
) := MP_IDLE;
END_TYPE

FUNCTION_BLOCK MaterialProportioningControl
VAR_INPUT
    estop : BOOL;
    opeMode : BOOL;
    valveAStart : BOOL;
    valveBStart : BOOL;
    valveCStart : BOOL;
    valveDStart : BOOL;
    mixMotorStart : BOOL;
    autoStart : BOOL;
    processMode : BOOL;
    levelSensor : INT;
    mixMotorComplete : BOOL;
END_VAR
VAR_OUTPUT
    valveARun : BOOL;
    valveBRun : BOOL;
    valveCRun : BOOL;
    valveDRun : BOOL;
    mixMotorRun : BOOL;
END_VAR
VAR
    tmp_trigValveA : R_TRIG;
    tmp_trigValveB : R_TRIG;
    tmp_trigValveC : R_TRIG;
    tmp_trigValveD : R_TRIG;
    tmp_trigMixMotor : R_TRIG;
    tmp_trigAutoStart : R_TRIG;

    manualValveARun : BOOL := FALSE;
    manualValveBRun : BOOL := FALSE;
    manualValveCRun : BOOL := FALSE;
    manualValveDRun : BOOL := FALSE;
    manualMixMotorRun : BOOL := FALSE;

    state : E_MaterialProportioningState := MP_IDLE;
    mixCompleteLatched : BOOL := FALSE;
END_VAR

tmp_trigValveA(CLK := valveAStart);
tmp_trigValveB(CLK := valveBStart);
tmp_trigValveC(CLK := valveCStart);
tmp_trigValveD(CLK := valveDStart);
tmp_trigMixMotor(CLK := mixMotorStart);
tmp_trigAutoStart(CLK := autoStart);

IF NOT estop THEN
    valveARun := FALSE;
    valveBRun := FALSE;
    valveCRun := FALSE;
    valveDRun := FALSE;
    mixMotorRun := FALSE;

ELSIF NOT opeMode THEN
    state := MP_IDLE;
    mixCompleteLatched := FALSE;

    IF tmp_trigValveA.Q THEN
        manualValveARun := NOT manualValveARun;
    END_IF;
    IF tmp_trigValveB.Q THEN
        manualValveBRun := NOT manualValveBRun;
    END_IF;
    IF tmp_trigValveC.Q THEN
        manualValveCRun := NOT manualValveCRun;
    END_IF;
    IF tmp_trigValveD.Q THEN
        manualValveDRun := NOT manualValveDRun;
    END_IF;
    IF tmp_trigMixMotor.Q THEN
        manualMixMotorRun := NOT manualMixMotorRun;
    END_IF;

    valveARun := manualValveARun;
    valveBRun := manualValveBRun;
    valveCRun := manualValveCRun;
    valveDRun := manualValveDRun;
    mixMotorRun := manualMixMotorRun;

ELSE
    IF tmp_trigAutoStart.Q THEN
        state := MP_FILL_A;
        mixCompleteLatched := FALSE;
    END_IF;

    CASE state OF
        MP_IDLE:
            valveARun := FALSE;
            valveBRun := FALSE;
            valveCRun := FALSE;
            valveDRun := FALSE;
            mixMotorRun := FALSE;

        MP_FILL_A:
            valveARun := TRUE;
            valveBRun := FALSE;
            valveCRun := FALSE;
            valveDRun := FALSE;
            mixMotorRun := FALSE;

            IF levelSensor >= 50 THEN
                valveARun := FALSE;
                valveBRun := TRUE;
                state := MP_FILL_B;
            END_IF;

        MP_FILL_B:
            valveARun := FALSE;
            valveBRun := TRUE;
            valveCRun := FALSE;
            valveDRun := FALSE;
            mixMotorRun := FALSE;

            IF levelSensor >= 80 THEN
                valveBRun := FALSE;
                IF NOT processMode THEN
                    mixMotorRun := TRUE;
                    mixCompleteLatched := FALSE;
                    state := MP_MIX_SIMPLE;
                ELSE
                    valveCRun := TRUE;
                    state := MP_FILL_C;
                END_IF;
            END_IF;

        MP_FILL_C:
            valveARun := FALSE;
            valveBRun := FALSE;
            valveCRun := TRUE;
            valveDRun := FALSE;
            mixMotorRun := FALSE;

            IF levelSensor >= 100 THEN
                valveCRun := FALSE;
                mixMotorRun := TRUE;
                mixCompleteLatched := FALSE;
                state := MP_MIX_C;
            END_IF;

        MP_MIX_SIMPLE:
            valveARun := FALSE;
            valveBRun := FALSE;
            valveCRun := FALSE;
            valveDRun := FALSE;
            mixMotorRun := TRUE;

            IF mixMotorComplete THEN
                mixCompleteLatched := TRUE;
            END_IF;

            IF mixCompleteLatched THEN
                mixMotorRun := FALSE;
                valveDRun := TRUE;
                state := MP_DONE;
            END_IF;

        MP_MIX_C:
            valveARun := FALSE;
            valveBRun := FALSE;
            valveCRun := FALSE;
            valveDRun := FALSE;
            mixMotorRun := TRUE;

            IF mixMotorComplete THEN
                mixCompleteLatched := TRUE;
            END_IF;

            IF mixCompleteLatched THEN
                mixMotorRun := FALSE;
                valveDRun := TRUE;
                state := MP_DONE;
            END_IF;

        MP_DONE:
            valveARun := FALSE;
            valveBRun := FALSE;
            valveCRun := FALSE;
            valveDRun := TRUE;
            mixMotorRun := FALSE;
    END_CASE;
END_IF;
END_FUNCTION_BLOCK

(* ---- public-hard-01.raw_candidate_02.st ---- *)
(* CONTRACT_RULES [] *)

(* ENGINEERING_CONTRACT
   - ESTOP: ESTOP=FALSE forces every output OFF in this scan; manual and auto commands are inhibited.
   - Manual runs: only while OpeMode=FALSE and ESTOP=TRUE; each start button rising edge toggles its retained output latch.
   - Auto sequence: AUTOSTART rising edge while OpeMode=TRUE enters FILL_A; output valves follow the sequence below.
   - Valve A: ON in FILL_A; Level>=50 closes A and opens B (PUB012).
   - Valve B: ON in FILL_B; Level>=80 closes B (PUB012/PUB013).
   - ProcessMode=FALSE: at Level>=80 mixer starts; MixMotorComplete latches completion, then mixer off and Valve D ON, sequence done (PUB014).
   - ProcessMode=TRUE: at Level>=80 Valve C opens; Level>=100 closes C and starts mixer; completion opens D (PUB014).
   - Mix complete is latched until the next AUTOSTART; Valve D remains ON in DONE because no stop/reset is stated.
   - Thresholds are inclusive >=; Level is INT cm; PROCESSMODE is read live at the 80 cm transition.
*)

TYPE E_MaterialProportioningState :
(
    MP_IDLE,
    MP_FILL_A,
    MP_FILL_B,
    MP_MIX_SIMPLE,
    MP_FILL_C,
    MP_MIX_C,
    MP_DONE
) := MP_IDLE;
END_TYPE;

FUNCTION_BLOCK MaterialProportioningControl
VAR_INPUT
    estop : BOOL;
    opeMode : BOOL;
    valveAStart : BOOL;
    valveBStart : BOOL;
    valveCStart : BOOL;
    valveDStart : BOOL;
    mixMotorStart : BOOL;
    autoStart : BOOL;
    processMode : BOOL;
    levelSensor : INT;
    mixMotorComplete : BOOL;
END_VAR
VAR_OUTPUT
    valveARun : BOOL;
    valveBRun : BOOL;
    valveCRun : BOOL;
    valveDRun : BOOL;
    mixMotorRun : BOOL;
END_VAR
VAR
    tmp_trigValveA : R_TRIG;
    tmp_trigValveB : R_TRIG;
    tmp_trigValveC : R_TRIG;
    tmp_trigValveD : R_TRIG;
    tmp_trigMixMotor : R_TRIG;
    tmp_trigAutoStart : R_TRIG;

    manualValveARun : BOOL := FALSE;
    manualValveBRun : BOOL := FALSE;
    manualValveCRun : BOOL := FALSE;
    manualValveDRun : BOOL := FALSE;
    manualMixMotorRun : BOOL := FALSE;

    state : E_MaterialProportioningState := MP_IDLE;
    mixCompleteLatched : BOOL := FALSE;
END_VAR

tmp_trigValveA(CLK := valveAStart);
tmp_trigValveB(CLK := valveBStart);
tmp_trigValveC(CLK := valveCStart);
tmp_trigValveD(CLK := valveDStart);
tmp_trigMixMotor(CLK := mixMotorStart);
tmp_trigAutoStart(CLK := autoStart);

IF NOT estop THEN
    valveARun := FALSE;
    valveBRun := FALSE;
    valveCRun := FALSE;
    valveDRun := FALSE;
    mixMotorRun := FALSE;

ELSIF NOT opeMode THEN
    state := MP_IDLE;
    mixCompleteLatched := FALSE;

    IF tmp_trigValveA.Q THEN
        manualValveARun := NOT manualValveARun;
    END_IF;
    IF tmp_trigValveB.Q THEN
        manualValveBRun := NOT manualValveBRun;
    END_IF;
    IF tmp_trigValveC.Q THEN
        manualValveCRun := NOT manualValveCRun;
    END_IF;
    IF tmp_trigValveD.Q THEN
        manualValveDRun := NOT manualValveDRun;
    END_IF;
    IF tmp_trigMixMotor.Q THEN
        manualMixMotorRun := NOT manualMixMotorRun;
    END_IF;

    valveARun := manualValveARun;
    valveBRun := manualValveBRun;
    valveCRun := manualValveCRun;
    valveDRun := manualValveDRun;
    mixMotorRun := manualMixMotorRun;

ELSE
    IF tmp_trigAutoStart.Q THEN
        state := MP_FILL_A;
        mixCompleteLatched := FALSE;
    END_IF;

    CASE state OF
        MP_IDLE:
            valveARun := FALSE;
            valveBRun := FALSE;
            valveCRun := FALSE;
            valveDRun := FALSE;
            mixMotorRun := FALSE;

        MP_FILL_A:
            valveARun := TRUE;
            valveBRun := FALSE;
            valveCRun := FALSE;
            valveDRun := FALSE;
            mixMotorRun := FALSE;

            IF levelSensor >= 50 THEN
                valveARun := FALSE;
                valveBRun := TRUE;
                state := MP_FILL_B;
            END_IF;

        MP_FILL_B:
            valveARun := FALSE;
            valveBRun := TRUE;
            valveCRun := FALSE;
            valveDRun := FALSE;
            mixMotorRun := FALSE;

            IF levelSensor >= 80 THEN
                valveBRun := FALSE;
                IF NOT processMode THEN
                    mixMotorRun := TRUE;
                    mixCompleteLatched := FALSE;
                    state := MP_MIX_SIMPLE;
                ELSE
                    IF levelSensor >= 100 THEN
                        valveCRun := FALSE;
                        mixMotorRun := TRUE;
                        mixCompleteLatched := FALSE;
                        state := MP_MIX_C;
                    ELSE
                        valveCRun := TRUE;
                        state := MP_FILL_C;
                    END_IF;
                END_IF;
            END_IF;

        MP_FILL_C:
            valveARun := FALSE;
            valveBRun := FALSE;
            valveCRun := TRUE;
            valveDRun := FALSE;
            mixMotorRun := FALSE;

            IF levelSensor >= 100 THEN
                valveCRun := FALSE;
                mixMotorRun := TRUE;
                mixCompleteLatched := FALSE;
                state := MP_MIX_C;
            END_IF;

        MP_MIX_SIMPLE:
            valveARun := FALSE;
            valveBRun := FALSE;
            valveCRun := FALSE;
            valveDRun := FALSE;
            mixMotorRun := TRUE;

            IF mixMotorComplete THEN
                mixCompleteLatched := TRUE;
            END_IF;

            IF mixCompleteLatched THEN
                mixMotorRun := FALSE;
                valveDRun := TRUE;
                state := MP_DONE;
            END_IF;

        MP_MIX_C:
            valveARun := FALSE;
            valveBRun := FALSE;
            valveCRun := FALSE;
            valveDRun := FALSE;
            mixMotorRun := TRUE;

            IF mixMotorComplete THEN
                mixCompleteLatched := TRUE;
            END_IF;

            IF mixCompleteLatched THEN
                mixMotorRun := FALSE;
                valveDRun := TRUE;
                state := MP_DONE;
            END_IF;

        MP_DONE:
            valveARun := FALSE;
            valveBRun := FALSE;
            valveCRun := FALSE;
            valveDRun := TRUE;
            mixMotorRun := FALSE;
    END_CASE;
END_IF;
END_FUNCTION_BLOCK
